                movel(spat_flatM_up_p, a=1.2, v=0.25, r=0.05)
                $ 2925 "Spatula_otw" "noBreak"
                movel(Spatula_otw_p, a=1.2, v=0.25)
                $ 2926 "switch_spat_F_M≔ False " "noBreak"
                global switch_spat_F_M=  False
              else:
                $ 2927 "ElseIf spatula≟'spatula_flat_S'" "noBreak"
                if (spatula == "spatula_flat_S"):
                  $ 2928 "MoveJ" "noBreak"
                  $ 2929 "Spatula_otw" "noBreak"
                  movej(get_inverse_kin(Spatula_otw_p, qnear=Spatula_otw_q), a=1.3962634015954636, v=1.0471975511965976)
                  $ 2930 "spat_flatS_up" "noBreak"
                  movej(get_inverse_kin(spat_flatS_up_p, qnear=spat_flatS_up_q), a=1.3962634015954636, v=1.0471975511965976, r=0.05)
                  $ 2931 "MoveL" "noBreak"
                  $ 2932 "spat_flatS_pick" "noBreak"
                  movel(spat_flatS_pick_p, a=1.2, v=0.25)
                  # begin: URCap Program Node
                  #   Source: Robotiq_Grippers, 3.17.0.105337, Robotiq Inc.
                  #   Type: Gripper
                  $ 2933 "Gripper Close (1)" "noBreak"
                  if not(gripper_connected[0]):
                    popup("Gripper 1 must be connected to run this program.", "No connection", False, True, True)
                  end
                  if not(rq_is_gripper_activated("1")):
                    popup("Gripper 1 is not activated. Go to Installation tab > Gripper to activate it and run the program again.", "Not activated", False, True, True)
                  end
                  rq_set_pos_spd_for(255, 0, 77, "1")
                  rq_wait_pos_spe_for_request(255, 0, 77, "1")
                  rq_go_to("1")
                  rq_wait("1")
                  # end: URCap Program Node
                  $ 2934 "spat_flatS_up" "noBreak"
                  movel(spat_flatS_up_p, a=1.2, v=0.25, r=0.05)
                  $ 2935 "Spatula_otw" "noBreak"
                  movel(Spatula_otw_p, a=1.2, v=0.25)
                  $ 2936 "switch_spat_F_S≔ False " "noBreak"
                  global switch_spat_F_S=  False
                end
              end
            end
          end
        end
        $ 2937 "weight_value≔get_weight()" "noBreak"
        global weight_value=get_weight()
        $ 2938 "auto_tilt_and_scoop(W_now, target_weight, weight_value)" "noBreak"
        auto_tilt_and_scoop(W_now, target_weight, weight_value)
        # begin: URCap Program Node
        #   Source: SensoPart VISOR Robotic, 2.0.6, SensoPart Industriesensorik GmbH
        #   Type: Approach Pose
        $ 2939 "Approach Pose" "noBreak"
        movej(pose_trans(easyPickPose,p[0.0000,0.0000,-0.0000,0.0000,0.0000,0.0000]),a=0.2618,v=0.1745,t=0.000000,r=0.000000)
        # end: URCap Program Node
        # begin: URCap Program Node
        #   Source: SensoPart VISOR Robotic, 2.0.6, SensoPart Industriesensorik GmbH
        #   Type: Target Pose
        $ 2940 "Target Pose" "noBreak"
        movel(pose_trans(easyPickPose,p[0.0000,0.0000,-0.0000,0.0000,0.0000,0.0000]),a=0.0500,v=0.0200,t=0.000000,r=0.000000)
        # end: URCap Program Node
        $ 2941 "Close Gripper" "noBreak"
        $ 2942 "dispense_pos≔get_actual_tcp_pose()" "noBreak"
        global dispense_pos= get_actual_tcp_pose ()
        $ 2943 "Loop weight_value≤target_weight" "noBreak"
        thread Thread_while_2943():
          while (True):
            $ 2944 "MoveL" "noBreak"
            $ 2945 "dispense_pos" "noBreak"
            movel(dispense_pos, a=0.2, v=0.1)
            $ 2946 "log_weight()" "noBreak"
            log_weight()
            $ 2947 "Wait: 0.5" "noBreak"
            sleep(0.5)
            $ 2948 "If level≥90.0" "noBreak"
            if (level >= 90.0):
              $ 2949 "Rotate()" "noBreak"
              Rotate()
            end
            $ 2950 "If level≤85" "noBreak"
            if (level <= 85):
              $ 2951 "tilt_to_home()" "noBreak"
              tilt_to_home()
            end
            $ 2952 "Wait: 0.5" "noBreak"
            sleep(0.5)
            $ 2953 "Start_thread≔ True " "noBreak"
            global Start_thread=  True
            $ 2954 "vib_thread≔ True " "noBreak"
            global vib_thread=  True
            $ 2956 "Wait: 0.5" "noBreak"
            sleep(0.5)
            $ 2962 "If diff ≥(target_g +(0.1*target_g))" "noBreak"
            if (diff  >= (target_g +(0.1*target_g))):
              $ 2963 "tilt_pose≔pose_trans(get_actual_tcp_pose(), p[0, 0, 0, 0, 0, 2.0])" "noBreak"
              global tilt_pose=pose_trans(get_actual_tcp_pose(), p[0, 0, 0, 0, 0, 2.0])
              $ 2964 "movel(tilt_pose, a=0.1, v=0.1, r=0.00001)" "noBreak"
              movel(tilt_pose, a=0.1, v=0.1, r=0.00001)
            else:
              $ 2965 "Else" "noBreak"
              $ 2966 "Loop weight_value≤target_weight and tilt_angle≥(-1.999) and tilt_angle≤0.5" "noBreak"
              thread Thread_while_2966():
                while (True):
                  $ 2967 "current_error≔target_weight-weight_value" "noBreak"
                  global current_error=target_weight-weight_value
                  $ 2968 "Integral_error≔Integral_error+current_error*dt" "noBreak"
                  global Integral_error=Integral_error+current_error*dt
                  $ 2969 "derivative≔(current_error-previous_error)/dt" "noBreak"
                  global derivative=(current_error-previous_error)/dt
                  $ 2970 "tilt_increment≔(kp*current_error)+(ki*Integral_error)+(kd*derivative)" "noBreak"
                  global tilt_increment=(kp*current_error)+(ki*Integral_error)+(kd*derivative)
                  $ 2971 "current_pose≔get_actual_tcp_pose()" "noBreak"
                  global current_pose= get_actual_tcp_pose ()
                  $ 2972 "tilt_angle≔current_pose[5]" "noBreak"
                  global tilt_angle=current_pose[5]
                  $ 2973 "tilt_pose≔pose_trans(current_pose, p[0, 0, 0, 0, 0, tilt_increment])" "noBreak"
                  global tilt_pose=pose_trans(current_pose, p[0, 0, 0, 0, 0, tilt_increment])
                  $ 2974 "movel(tilt_pose, a=0.1, v=0.1, r=0.00001)" "noBreak"
                  movel(tilt_pose, a=0.1, v=0.1, r=0.00001)
                  $ 2975 "previous_error≔current_error" "noBreak"
                  global previous_error=current_error
                end
              end
              if (weight_value <= target_weight  and  tilt_angle >= (-1.999)  and  tilt_angle <= 0.5):
                global thread_handler_2966=run Thread_while_2966()
                while (weight_value <= target_weight  and  tilt_angle >= (-1.999)  and  tilt_angle <= 0.5):
                  sync()
                end
                kill thread_handler_2966
              end
            end
            $ 2976 "Start_thread≔ False " "noBreak"
            global Start_thread=  False
            $ 2978 "weight_value≔get_weight()" "noBreak"
            global weight_value=get_weight()
            $ 2979 "tilt_angle≔-1" "noBreak"
            global tilt_angle=-1
            $ 2980 "Wait: 0.5" "noBreak"
            sleep(0.5)
            $ 2981 "vib_thread≔ False " "noBreak"
            global vib_thread=  False
            $ 2982 "MoveL" "noBreak"
            $ 2983 "dispense_pos" "noBreak"
            movel(dispense_pos, a=0.5, v=0.25)
            $ 2984 "compute_level_percent(W_now, weight_value)" "noBreak"
            compute_level_percent(W_now, weight_value)
            $ 2985 "send_level_info()" "noBreak"
            send_level_info()
            $ 2987 "spatula≔select_spatula(Flowability,level,diff,density)" "noBreak"
            global spatula=select_spatula(Flowability,level,diff,density)
            $ 2989 "Wait: 0.2" "noBreak"
            sleep(0.2)
            $ 2991 "Integral_error≔0" "noBreak"
            global Integral_error=0
            $ 2992 "current_error≔0" "noBreak"
            global current_error=0
            $ 2993 "previous_error≔0" "noBreak"
            global previous_error=0
            $ 2994 "Set AO[0]=0.0" "noBreak"
            set_standard_analog_out(0, 0.0)
            $ 2995 "Wait: 0.2" "noBreak"
            sleep(0.2)
            $ 2996 "send_spatula_info()" "noBreak"
            send_spatula_info()
            $ 2997 "If spatula ≟ 'spatula_M' and switch_spat_M≟ True " "noBreak"
            if (spatula  ==  "spatula_M"  and  switch_spat_M ==   True  ):
              $ 2998 "MoveJ" "noBreak"
              $ 2999 "Spatula_otw" "noBreak"
              movej(get_inverse_kin(Spatula_otw_p, qnear=Spatula_otw_q), a=1.3962634015954636, v=1.0471975511965976)
              $ 3000 "spat_L_up" "noBreak"
              movej(get_inverse_kin(spat_L_up_p, qnear=spat_L_up_q), a=1.3962634015954636, v=1.0471975511965976)
              $ 3001 "MoveL" "noBreak"
              $ 3002 "spat_L_side" "noBreak"
              movel(spat_L_side_p, a=1.2, v=0.25)
              $ 3003 "spat_L_lift" "noBreak"
              movel(spat_L_lift_p, a=1.2, v=0.25)
              $ 3004 "spat_L_pick" "noBreak"
              movel(spat_L_pick_p, a=1.2, v=0.25)
              # begin: URCap Program Node
              #   Source: Robotiq_Grippers, 3.17.0.105337, Robotiq Inc.
              #   Type: Gripper
              $ 3005 "Gripper Open (1)" "noBreak"
              if not(gripper_connected[0]):
                popup("Gripper 1 must be connected to run this program.", "No connection", False, True, True)
              end
              if not(rq_is_gripper_activated("1")):
                popup("Gripper 1 is not activated. Go to Installation tab > Gripper to activate it and run the program again.", "Not activated", False, True, True)
              end
              rq_set_pos_spd_for(0, 255, 77, "1")
              rq_wait_pos_spe_for_request(0, 255, 77, "1")
              rq_go_to("1")
              rq_wait("1")
              # end: URCap Program Node
              $ 3006 "spat_M_pick" "noBreak"
              movel(spat_M_pick_p, a=1.2, v=0.25)
              # begin: URCap Program Node
              #   Source: Robotiq_Grippers, 3.17.0.105337, Robotiq Inc.
              #   Type: Gripper
              $ 3007 "Gripper Close (1)" "noBreak"
              if not(gripper_connected[0]):
                popup("Gripper 1 must be connected to run this program.", "No connection", False, True, True)
              end
              if not(rq_is_gripper_activated("1")):
                popup("Gripper 1 is not activated. Go to Installation tab > Gripper to activate it and run the program again.", "Not activated", False, True, True)
              end
              rq_set_pos_spd_for(255, 0, 77, "1")
              rq_wait_pos_spe_for_request(255, 0, 77, "1")
              rq_go_to("1")
              rq_wait("1")
              # end: URCap Program Node
              $ 3008 "spat_M_up" "noBreak"
              movel(spat_M_up_p, a=1.2, v=0.25)
              $ 3009 "Spatula_otw" "noBreak"
              movel(Spatula_otw_p, a=1.2, v=0.25)
              $ 3010 "switch_spat_M≔ False " "noBreak"
              global switch_spat_M=  False
            else:
              $ 3011 "ElseIf spatula ≟ 'spatula_S' and switch_spat_S ≟ True " "noBreak"
              if (spatula  ==  "spatula_S" and switch_spat_S  ==   True  ):
                $ 3012 "MoveL" "noBreak"
                $ 3013 "Spatula_otw" "noBreak"
                movel(Spatula_otw_p, a=1.2, v=0.25)
                $ 3014 "spat_M_up" "noBreak"
                movel(spat_M_up_p, a=1.2, v=0.25)
                $ 3015 "spat_M_pick" "noBreak"
                movel(spat_M_pick_p, a=1.2, v=0.25)
                # begin: URCap Program Node
                #   Source: Robotiq_Grippers, 3.17.0.105337, Robotiq Inc.
                #   Type: Gripper
                $ 3016 "Gripper Open (1)" "noBreak"
                if not(gripper_connected[0]):
                  popup("Gripper 1 must be connected to run this program.", "No connection", False, True, True)
                end
                if not(rq_is_gripper_activated("1")):
                  popup("Gripper 1 is not activated. Go to Installation tab > Gripper to activate it and run the program again.", "Not activated", False, True, True)
                end
                rq_set_pos_spd_for(0, 255, 77, "1")
                rq_wait_pos_spe_for_request(0, 255, 77, "1")
                rq_go_to("1")
                rq_wait("1")
                # end: URCap Program Node
                $ 3017 "spat_S_pick" "noBreak"
                movel(spat_S_pick_p, a=1.2, v=0.25)
                # begin: URCap Program Node
                #   Source: Robotiq_Grippers, 3.17.0.105337, Robotiq Inc.
                #   Type: Gripper
                $ 3018 "Gripper Close (1)" "noBreak"
                if not(gripper_connected[0]):
                  popup("Gripper 1 must be connected to run this program.", "No connection", False, True, True)
                end
                if not(rq_is_gripper_activated("1")):
                  popup("Gripper 1 is not activated. Go to Installation tab > Gripper to activate it and run the program again.", "Not activated", False, True, True)
                end
                rq_set_pos_spd_for(255, 0, 77, "1")
                rq_wait_pos_spe_for_request(255, 0, 77, "1")
                rq_go_to("1")
                rq_wait("1")
                # end: URCap Program Node
                $ 3019 "spat_S_up" "noBreak"
                movel(spat_S_up_p, a=1.2, v=0.25)
                $ 3020 "Spatula_otw" "noBreak"
                movel(Spatula_otw_p, a=1.2, v=0.25)
                $ 3021 "switch_spat_S≔ False " "noBreak"
                global switch_spat_S=  False
              else:
                $ 3022 "ElseIf spatula≟'spatula_flat_S'  and switch_spat_F_S ≟ True " "noBreak"
                if (spatula == "spatula_flat_S"   and  switch_spat_F_S  ==   True  ):
                  $ 3023 "MoveL" "noBreak"
                  $ 3024 "Spatula_otw" "noBreak"
                  movel(Spatula_otw_p, a=1.2, v=0.25)
                  $ 3025 "spat_flatM_up" "noBreak"
                  movel(spat_flatM_up_p, a=1.2, v=0.25)
                  $ 3026 "spat_flatM_pick" "noBreak"
                  movel(spat_flatM_pick_p, a=1.2, v=0.25)
                  # begin: URCap Program Node
                  #   Source: Robotiq_Grippers, 3.17.0.105337, Robotiq Inc.
                  #   Type: Gripper
                  $ 3027 "Gripper Open (1)" "noBreak"
                  if not(gripper_connected[0]):
                    popup("Gripper 1 must be connected to run this program.", "No connection", False, True, True)
                  end
                  if not(rq_is_gripper_activated("1")):
                    popup("Gripper 1 is not activated. Go to Installation tab > Gripper to activate it and run the program again.", "Not activated", False, True, True)
                  end
                  rq_set_pos_spd_for(0, 0, 77, "1")
                  rq_wait_pos_spe_for_request(0, 0, 77, "1")
                  rq_go_to("1")
                  rq_wait("1")
                  # end: URCap Program Node
                  $ 3028 "spat_flatS_pick" "noBreak"
                  movel(spat_flatS_pick_p, a=1.2, v=0.25)
                  # begin: URCap Program Node
                  #   Source: Robotiq_Grippers, 3.17.0.105337, Robotiq Inc.
                  #   Type: Gripper
                  $ 3029 "Gripper Close (1)" "noBreak"
                  if not(gripper_connected[0]):
                    popup("Gripper 1 must be connected to run this program.", "No connection", False, True, True)
                  end
                  if not(rq_is_gripper_activated("1")):
                    popup("Gripper 1 is not activated. Go to Installation tab > Gripper to activate it and run the program again.", "Not activated", False, True, True)
                  end
                  rq_set_pos_spd_for(255, 0, 77, "1")
                  rq_wait_pos_spe_for_request(255, 0, 77, "1")
                  rq_go_to("1")
                  rq_wait("1")
                  # end: URCap Program Node
                  $ 3030 "spat_flatS_up" "noBreak"
                  movel(spat_flatS_up_p, a=1.2, v=0.25)
                  $ 3031 "Spatula_otw" "noBreak"
                  movel(Spatula_otw_p, a=1.2, v=0.25)
                  $ 3032 "switch_spat_F_S≔ False " "noBreak"
                  global switch_spat_F_S=  False
                end
              end
            end
            $ 3033 "auto_tilt_and_scoop(W_now, target_weight, weight_value)" "noBreak"
            auto_tilt_and_scoop(W_now, target_weight, weight_value)
            $ 3034 "Wait: 0.5" "noBreak"
            sleep(0.5)
          end
        end
        if (weight_value <= target_weight):
          global thread_handler_2943=run Thread_while_2943()
          while (weight_value <= target_weight):
            sync()
          end
          kill thread_handler_2943
        end
        $ 3035 "Start_thread≔ False " "noBreak"
        global Start_thread=  False
        $ 3036 "Wait: 0.5" "noBreak"
        sleep(0.5)
        $ 3037 "vib_thread≔ False " "noBreak"
        global vib_thread=  False
        # begin: URCap Program Node
        #   Source: SensoPart VISOR Robotic, 2.0.6, SensoPart Industriesensorik GmbH
        #   Type: Exit Pose
        $ 3039 "Exit Pose" "noBreak"
        movel(pose_trans(easyPickPose,p[0.0000,0.0000,-0.0000,0.0000,0.0000,0.0000]),a=0.5000,v=0.2500,t=0.000000,r=0.000000)
        # end: URCap Program Node
        easyPickObjTaken = True
      end
      # end: URCap Program Node
      # begin: URCap Program Node
      #   Source: SensoPart VISOR Robotic, 2.0.6, SensoPart Industriesensorik GmbH
      #   Type: No Object Detected
      $ 3040 "No Object Detected" "noBreak"
      if (visor_partsFound(easyPickVisorId) < 1):
        $ 3041 "Popup: No weigh scale detected" "noBreak"
        popup("No weigh scale detected", "Message", False, False, blocking=True)
        else:
      end
      # end: URCap Program Node
    end
    easyPickCount_4 = easyPickCount_4 + 1
    visor_easyPickUpdate(easyPickVisorId, "counter", easyPickCount_4)
    visor_easyPickSetIdent("6c09fd", easyPickVisorId)
    # end: URCap Program Node
  end
  visorFuncEasyPick_ff2f00()
  # end: URCap Program Node
  $ 3044 "MoveJ"
  $ 3045 "dispense_pos" "breakAfter"
  movej(dispense_pos, a=0.5235987755982988, v=0.4363323129985824)
  $ 3046 "after_scoop()"
  after_scoop()
  $ 3047 "Place spatula back to the rack"
  $ 3048 "If spatula≟'spatula_M'"
  if (spatula == "spatula_M"):
    $ 3049 "MoveJ"
    $ 3050 "Spatula_otw" "breakAfter"
    movej(get_inverse_kin(Spatula_otw_p, qnear=Spatula_otw_q), a=1.3962634015954636, v=1.0471975511965976)
    $ 3051 "spat_M_up" "breakAfter"
    movej(get_inverse_kin(spat_M_up_p, qnear=spat_M_up_q), a=1.3962634015954636, v=1.0471975511965976)
    $ 3052 "MoveL"
    $ 3053 "spat_M_pick" "breakAfter"
    movel(spat_M_pick_p, a=1.2, v=0.25)
    # begin: URCap Program Node
    #   Source: Robotiq_Grippers, 3.17.0.105337, Robotiq Inc.
    #   Type: Gripper
    $ 3054 "Gripper Open (1)"
    if not(gripper_connected[0]):
      popup("Gripper 1 must be connected to run this program.", "No connection", False, True, True)
    end
    if not(rq_is_gripper_activated("1")):
      popup("Gripper 1 is not activated. Go to Installation tab > Gripper to activate it and run the program again.", "Not activated", False, True, True)
    end
    rq_set_pos_spd_for(0, 128, 77, "1")
    rq_wait_pos_spe_for_request(0, 128, 77, "1")
    rq_go_to("1")
    rq_wait("1")
    # end: URCap Program Node
    $ 3055 "spat_M_up" "breakAfter"
    movel(spat_M_up_p, a=1.2, v=0.25)
    $ 3056 "Home (Safe)"
    movej([-1.2302089344500047, -1.2969853503591224, -1.875639182904262, -1.539621866126728, 1.5731943360401213, -2.80099559440227], a=1.3962634015954636, v=1.0471975511965976)
  else:
    $ 3057 "ElseIf spatula≟'spatula_flat_S'"
    if (spatula == "spatula_flat_S"):
      $ 3058 "MoveJ"
      $ 3059 "Spatula_otw" "breakAfter"
      movej(get_inverse_kin(Spatula_otw_p, qnear=Spatula_otw_q), a=1.3962634015954636, v=1.0471975511965976)
      $ 3060 "spat_flatS_up" "breakAfter"
      movej(get_inverse_kin(spat_flatS_up_p, qnear=spat_flatS_up_q), a=1.3962634015954636, v=1.0471975511965976)
      $ 3061 "MoveL"
      $ 3062 "spat_flatS_pick" "breakAfter"
      movel(spat_flatS_pick_p, a=1.2, v=0.25)
      # begin: URCap Program Node
      #   Source: Robotiq_Grippers, 3.17.0.105337, Robotiq Inc.
      #   Type: Gripper
      $ 3063 "Gripper Open (1)"
      if not(gripper_connected[0]):
        popup("Gripper 1 must be connected to run this program.", "No connection", False, True, True)
      end
      if not(rq_is_gripper_activated("1")):
        popup("Gripper 1 is not activated. Go to Installation tab > Gripper to activate it and run the program again.", "Not activated", False, True, True)
      end
      rq_set_pos_spd_for(0, 128, 77, "1")
      rq_wait_pos_spe_for_request(0, 128, 77, "1")
      rq_go_to("1")
      rq_wait("1")
      # end: URCap Program Node
      $ 3064 "spat_flatS_up" "breakAfter"
      movel(spat_flatS_up_p, a=1.2, v=0.25)
      $ 3065 "Home (Safe)"
      movej([-1.2302089344500047, -1.2969853503591224, -1.875639182904262, -1.539621866126728, 1.5731943360401213, -2.80099559440227], a=1.3962634015954636, v=1.0471975511965976)
    end
  end
  $ 3066 "Pick container from PoTS"
  $ 3067 "cont_place_offs≔pose_add(container_place, p[0.05,0,0,0,0,0])"
  global cont_place_offs=pose_add(container_place, p[0.05,0,0,0,0,0])
  $ 3068 "MoveJ"
  $ 3069 "cont_place_offs" "breakAfter"
  movej(cont_place_offs, a=1.3962634015954636, v=1.0471975511965976)
  $ 3070 "container_place" "breakAfter"
  movej(container_place, a=1.3962634015954636, v=1.0471975511965976)
  $ 3071 "MoveL"
  $ 3072 "target_pose" "breakAfter"
  movel(target_pose, a=1.2, v=0.25)
  # begin: URCap Program Node
  #   Source: Robotiq_Grippers, 3.17.0.105337, Robotiq Inc.
  #   Type: Gripper
  $ 3073 "Gripper Close (1)"
  if not(gripper_connected[0]):
    popup("Gripper 1 must be connected to run this program.", "No connection", False, True, True)
  end
  if not(rq_is_gripper_activated("1")):
    popup("Gripper 1 is not activated. Go to Installation tab > Gripper to activate it and run the program again.", "Not activated", False, True, True)
  end
  rq_set_pos_spd_for(255, 77, 77, "1")
  rq_wait_pos_spe_for_request(255, 77, 77, "1")
  rq_go_to("1")
  rq_wait("1")
  # end: URCap Program Node
  $ 3074 "container_place" "breakAfter"
  movel(container_place, a=0.6, v=0.1)
  $ 3075 "powder_position≔'Position1'"
  global powder_position="Position1"
  $ 3076 "Place Powder container back to holder"
  $ 3077 "If powder_position ≟ 'Position1'"
  if (powder_position  ==  "Position1"):
    $ 3078 "MoveL"
    $ 3079 "Postions_otw" "breakAfter"
    movel(Postions_otw_p, a=1.2, v=0.25, r=0.01)
    $ 3080 "MoveL"
    $ 3081 "PosA_up" "breakAfter"
    movel(PosA_up_p, a=1.2, v=0.25)
    $ 3082 "PosA_pick" "breakAfter"
    movel(PosA_pick_p, a=0.3, v=0.05)
    # begin: URCap Program Node
    #   Source: Robotiq_Grippers, 3.17.0.105337, Robotiq Inc.
    #   Type: Gripper
    $ 3083 "Gripper Open (1)"
    if not(gripper_connected[0]):
      popup("Gripper 1 must be connected to run this program.", "No connection", False, True, True)
    end
    if not(rq_is_gripper_activated("1")):
      popup("Gripper 1 is not activated. Go to Installation tab > Gripper to activate it and run the program again.", "Not activated", False, True, True)
    end
    rq_set_pos_spd_for(0, 128, 77, "1")
    rq_wait_pos_spe_for_request(0, 128, 77, "1")
    rq_go_to("1")
    rq_wait("1")
    # end: URCap Program Node
    $ 3084 "PosA_up" "breakAfter"
    movel(PosA_up_p, a=1.2, v=0.25)
    $ 3085 "Postions_otw" "breakAfter"
    movel(Postions_otw_p, a=1.2, v=0.25, r=0.05)
  else:
    $ 3086 "ElseIf powder_position≟'Position2'"
    if (powder_position == "Position2"):
      $ 3087 "MoveL"
      $ 3088 "Postions_otw" "breakAfter"
      movel(Postions_otw_p, a=1.2, v=0.25, r=0.01)
      $ 3089 "MoveL"
      $ 3090 "PosB_up" "breakAfter"
      movel(PosB_up_p, a=1.2, v=0.25, r=0.01)
      $ 3091 "PosB_pick" "breakAfter"
      movel(PosB_pick_p, a=0.3, v=0.05)
      # begin: URCap Program Node
      #   Source: Robotiq_Grippers, 3.17.0.105337, Robotiq Inc.
      #   Type: Gripper
      $ 3092 "Gripper Open (1)"
      if not(gripper_connected[0]):
        popup("Gripper 1 must be connected to run this program.", "No connection", False, True, True)
      end
      if not(rq_is_gripper_activated("1")):
        popup("Gripper 1 is not activated. Go to Installation tab > Gripper to activate it and run the program again.", "Not activated", False, True, True)
      end
      rq_set_pos_spd_for(0, 128, 77, "1")
      rq_wait_pos_spe_for_request(0, 128, 77, "1")
      rq_go_to("1")
      rq_wait("1")
      # end: URCap Program Node
      $ 3093 "PosB_up" "breakAfter"
      movel(PosB_up_p, a=1.2, v=0.25)
      $ 3094 "Postions_otw" "breakAfter"
      movel(Postions_otw_p, a=1.2, v=0.25, r=0.05)
    else:
      $ 3095 "ElseIf powder_position≟'Position3'"
      if (powder_position == "Position3"):
        $ 3096 "MoveL"
        $ 3097 "Postions_otw" "breakAfter"
        movel(Postions_otw_p, a=1.2, v=0.25, r=0.01)
        $ 3098 "MoveL"
        $ 3099 "PosC_up" "breakAfter"
        movel(PosC_up_p, a=1.2, v=0.25, r=0.01)
        $ 3100 "PosC_pick" "breakAfter"
        movel(PosC_pick_p, a=0.3, v=0.05)
        # begin: URCap Program Node
        #   Source: Robotiq_Grippers, 3.17.0.105337, Robotiq Inc.
        #   Type: Gripper
        $ 3101 "Gripper Open (1)"
        if not(gripper_connected[0]):
          popup("Gripper 1 must be connected to run this program.", "No connection", False, True, True)
        end
        if not(rq_is_gripper_activated("1")):
          popup("Gripper 1 is not activated. Go to Installation tab > Gripper to activate it and run the program again.", "Not activated", False, True, True)
        end
        rq_set_pos_spd_for(0, 128, 77, "1")
        rq_wait_pos_spe_for_request(0, 128, 77, "1")
        rq_go_to("1")
        rq_wait("1")
        # end: URCap Program Node
        $ 3102 "PosC_up" "breakAfter"
        movel(PosC_up_p, a=1.2, v=0.25)
        $ 3103 "Postions_otw" "breakAfter"
        movel(Postions_otw_p, a=1.2, v=0.25, r=0.05)
      end
    end
  end
  $ 3104 "Cap the container"
  $ 3105 "If powder_position ≟ 'Position1'"
  if (powder_position  ==  "Position1"):
    $ 3106 "MoveJ"
    $ 3107 "Cap_Pos1_up" "breakAfter"
    movej(get_inverse_kin(Cap_Pos1_up_p, qnear=Cap_Pos1_up_q), a=1.3962634015954636, v=1.0471975511965976)
    $ 3108 "MoveL"
    $ 3109 "Cap_pos1" "breakAfter"
    movel(Cap_pos1_p, a=0.3, v=0.05)
  else:
    $ 3110 "ElseIf powder_position≟'Position2'"
    if (powder_position == "Position2"):
      $ 3111 "MoveJ"
      $ 3112 "Cap_Pos2_up" "breakAfter"
      movej(get_inverse_kin(Cap_Pos2_up_p, qnear=Cap_Pos2_up_q), a=1.3962634015954636, v=1.0471975511965976)
      $ 3113 "MoveL"
      $ 3114 "Cap_Pos2" "breakAfter"
      movel(Cap_Pos2_p, a=0.3, v=0.05)
    else:
      $ 3115 "ElseIf powder_position≟'Position3'"
      if (powder_position == "Position3"):
        $ 3116 "MoveJ"
        $ 3117 "Cap_Pos3_up" "breakAfter"
        movej(get_inverse_kin(Cap_Pos3_up_p, qnear=Cap_Pos3_up_q), a=1.3962634015954636, v=1.0471975511965976)
        $ 3118 "MoveL"
        $ 3119 "Cap_pos3" "breakAfter"
        movel(Cap_pos3_p, a=0.3, v=0.05)
      end
    end
  end
  $ 3120 "Capping motion"
  # begin: URCap Program Node
  #   Source: Robotiq_Grippers, 3.17.0.105337, Robotiq Inc.
  #   Type: Gripper
  $ 3121 "Gripper Move30mm (1)"
  if not(gripper_connected[0]):
    popup("Gripper 1 must be connected to run this program.", "No connection", False, True, True)
  end
  if not(rq_is_gripper_activated("1")):
    popup("Gripper 1 is not activated. Go to Installation tab > Gripper to activate it and run the program again.", "Not activated", False, True, True)
  end
  rq_set_pos_spd_for(110, 77, 77, "1")
  rq_wait_pos_spe_for_request(110, 77, 77, "1")
  rq_go_to("1")
  rq_wait("1")
  # end: URCap Program Node
  $ 3122 "Loop 2 times"
  Loop_4 = 0
  while (Loop_4 < 2):
    $ 3128 "Cap_CW≔pose_add(get_actual_tcp_pose(), p[0,0,0,0,0,2.2])"
    global Cap_CW= pose_add ( get_actual_tcp_pose (), p[0,0,0,0,0,2.2])
    $ 3129 "MoveL"
    $ 3130 "Cap_CW" "breakAfter"
    movel(Cap_CW, a=1.2, v=0.25)
    # begin: URCap Program Node
    #   Source: Robotiq_Grippers, 3.17.0.105337, Robotiq Inc.
    #   Type: Gripper
    $ 3131 "Gripper Move25mm (1)"
    if not(gripper_connected[0]):
      popup("Gripper 1 must be connected to run this program.", "No connection", False, True, True)
    end
    if not(rq_is_gripper_activated("1")):
      popup("Gripper 1 is not activated. Go to Installation tab > Gripper to activate it and run the program again.", "Not activated", False, True, True)
    end
    rq_set_pos_spd_for(133, 77, 77, "1")
    rq_wait_pos_spe_for_request(133, 77, 77, "1")
    rq_go_to("1")
    rq_wait("1")
    # end: URCap Program Node
    $ 3132 "Cap_CCW≔pose_add(get_actual_tcp_pose(), p[0,0,0,0,0,-2.2])"
    global Cap_CCW= pose_add ( get_actual_tcp_pose (), p[0,0,0,0,0,-2.2])
    $ 3133 "MoveL"
    $ 3134 "Cap_CCW" "breakAfter"
    movel(Cap_CCW, a=1.2, v=0.25)
    # begin: URCap Program Node
    #   Source: Robotiq_Grippers, 3.17.0.105337, Robotiq Inc.
    #   Type: Gripper
    $ 3135 "Gripper Move30mm (1)"
    if not(gripper_connected[0]):
      popup("Gripper 1 must be connected to run this program.", "No connection", False, True, True)
    end
    if not(rq_is_gripper_activated("1")):
      popup("Gripper 1 is not activated. Go to Installation tab > Gripper to activate it and run the program again.", "Not activated", False, True, True)
    end
    rq_set_pos_spd_for(110, 77, 77, "1")
    rq_wait_pos_spe_for_request(110, 77, 77, "1")
    rq_go_to("1")
    rq_wait("1")
    # end: URCap Program Node
    Loop_4 = Loop_4 + 1
  end
  # begin: URCap Program Node
  #   Source: Robotiq_Grippers, 3.17.0.105337, Robotiq Inc.
  #   Type: Gripper
  $ 3136 "Gripper Open (1)"
  if not(gripper_connected[0]):
    popup("Gripper 1 must be connected to run this program.", "No connection", False, True, True)
  end
  if not(rq_is_gripper_activated("1")):
    popup("Gripper 1 is not activated. Go to Installation tab > Gripper to activate it and run the program again.", "Not activated", False, True, True)
  end
  rq_set_pos_spd_for(0, 77, 77, "1")
  rq_wait_pos_spe_for_request(0, 77, 77, "1")
  rq_go_to("1")
  rq_wait("1")
  # end: URCap Program Node
  $ 3137 "after_capping≔pose_add(get_actual_tcp_pose(), p[0,0,0.05,0,0,0])"
  global after_capping=pose_add(get_actual_tcp_pose(), p[0,0,0.05,0,0,0])
  $ 3138 "MoveL"
  $ 3139 "after_capping" "breakAfter"
  movel(after_capping, a=1.2, v=0.25)
  $ 3140 "Home (Safe)"
  movej([-1.2302089344500047, -1.2969853503591224, -1.875639182904262, -1.539621866126728, 1.5731943360401213, -2.80099559440227], a=1.3962634015954636, v=1.0471975511965976)
  elif (44 == switch_1):
    $ 3203 "Case 44"
    $ 3204 "Decap Container for recipe"
    $ 3206 "If powder_position ≟ 'Position1'"
    if (powder_position  ==  "Position1"):
      $ 3207 "MoveJ"
      $ 3208 "Postions_otw" "breakAfter"
      movej(get_inverse_kin(Postions_otw_p, qnear=Postions_otw_q), a=1.3962634015954636, v=1.0471975511965976, r=0.01)
      # begin: URCap Program Node
      #   Source: Robotiq_Grippers, 3.17.0.105337, Robotiq Inc.
      #   Type: Gripper
      $ 3209 "Gripper Open (1)"
      if not(gripper_connected[0]):
        popup("Gripper 1 must be connected to run this program.", "No connection", False, True, True)
      end
      if not(rq_is_gripper_activated("1")):
        popup("Gripper 1 is not activated. Go to Installation tab > Gripper to activate it and run the program again.", "Not activated", False, True, True)
      end
      rq_set_pos_spd_for(0, 127, 77, "1")
      rq_wait_pos_spe_for_request(0, 127, 77, "1")
      rq_go_to("1")
      rq_wait("1")
      # end: URCap Program Node
      $ 3210 "MoveL"
      $ 3211 "PosA_up" "breakAfter"
      movel(PosA_up_p, a=1.2, v=0.25)
      $ 3212 "PosA_pick" "breakAfter"
      movel(PosA_pick_p, a=1.2, v=0.25)
      # begin: URCap Program Node
      #   Source: Robotiq_Grippers, 3.17.0.105337, Robotiq Inc.
      #   Type: Gripper
      $ 3213 "Gripper Close (1)"
      if not(gripper_connected[0]):
        popup("Gripper 1 must be connected to run this program.", "No connection", False, True, True)
      end
      if not(rq_is_gripper_activated("1")):
        popup("Gripper 1 is not activated. Go to Installation tab > Gripper to activate it and run the program again.", "Not activated", False, True, True)
      end
      rq_set_pos_spd_for(255, 127, 77, "1")
      rq_wait_pos_spe_for_request(255, 127, 77, "1")
      rq_go_to("1")
      rq_wait("1")
      # end: URCap Program Node
      $ 3214 "PosA_up" "breakAfter"
      movel(PosA_up_p, a=0.3, v=0.04)
      $ 3215 "Postions_otw" "breakAfter"
      movel(Postions_otw_p, a=1.2, v=0.25, r=0.01)
    else:
      $ 3216 "ElseIf powder_position≟'Position2'"
      if (powder_position == "Position2"):
        $ 3217 "MoveJ"
        $ 3218 "Postions_otw" "breakAfter"
        movej(get_inverse_kin(Postions_otw_p, qnear=Postions_otw_q), a=1.3962634015954636, v=1.0471975511965976, r=0.01)
        # begin: URCap Program Node
        #   Source: Robotiq_Grippers, 3.17.0.105337, Robotiq Inc.
        #   Type: Gripper
        $ 3219 "Gripper Open (1)"
        if not(gripper_connected[0]):
          popup("Gripper 1 must be connected to run this program.", "No connection", False, True, True)
        end
        if not(rq_is_gripper_activated("1")):
          popup("Gripper 1 is not activated. Go to Installation tab > Gripper to activate it and run the program again.", "Not activated", False, True, True)
        end
        rq_set_pos_spd_for(0, 127, 77, "1")
        rq_wait_pos_spe_for_request(0, 127, 77, "1")
        rq_go_to("1")
        rq_wait("1")
        # end: URCap Program Node
        $ 3220 "MoveL"
        $ 3221 "PosB_up" "breakAfter"
        movel(PosB_up_p, a=1.2, v=0.25, r=0.01)
        $ 3222 "PosB_pick" "breakAfter"
        movel(PosB_pick_p, a=1.2, v=0.25)
        # begin: URCap Program Node
        #   Source: Robotiq_Grippers, 3.17.0.105337, Robotiq Inc.
        #   Type: Gripper
        $ 3223 "Gripper Close (1)"
        if not(gripper_connected[0]):
          popup("Gripper 1 must be connected to run this program.", "No connection", False, True, True)
        end
        if not(rq_is_gripper_activated("1")):
          popup("Gripper 1 is not activated. Go to Installation tab > Gripper to activate it and run the program again.", "Not activated", False, True, True)
        end
        rq_set_pos_spd_for(255, 127, 77, "1")
        rq_wait_pos_spe_for_request(255, 127, 77, "1")
        rq_go_to("1")
        rq_wait("1")
        # end: URCap Program Node
        $ 3224 "PosB_up" "breakAfter"
        movel(PosB_up_p, a=0.4, v=0.05)
        $ 3225 "Postions_otw" "breakAfter"
        movel(Postions_otw_p, a=1.2, v=0.25)
      else:
        $ 3226 "ElseIf powder_position≟'Position3'"
        if (powder_position == "Position3"):
          $ 3227 "MoveJ"
          $ 3228 "Postions_otw" "breakAfter"
          movej(get_inverse_kin(Postions_otw_p, qnear=Postions_otw_q), a=1.3962634015954636, v=1.0471975511965976, r=0.01)
          # begin: URCap Program Node
          #   Source: Robotiq_Grippers, 3.17.0.105337, Robotiq Inc.
          #   Type: Gripper
          $ 3229 "Gripper Open (1)"
          if not(gripper_connected[0]):
            popup("Gripper 1 must be connected to run this program.", "No connection", False, True, True)
          end
          if not(rq_is_gripper_activated("1")):
            popup("Gripper 1 is not activated. Go to Installation tab > Gripper to activate it and run the program again.", "Not activated", False, True, True)
          end
          rq_set_pos_spd_for(0, 127, 77, "1")
          rq_wait_pos_spe_for_request(0, 127, 77, "1")
          rq_go_to("1")
          rq_wait("1")
          # end: URCap Program Node
          $ 3230 "MoveL"
          $ 3231 "PosC_up" "breakAfter"
          movel(PosC_up_p, a=1.2, v=0.25, r=0.01)
          $ 3232 "PosC_pick" "breakAfter"
          movel(PosC_pick_p, a=1.2, v=0.25)
          # begin: URCap Program Node
          #   Source: Robotiq_Grippers, 3.17.0.105337, Robotiq Inc.
          #   Type: Gripper
          $ 3233 "Gripper Close (1)"
          if not(gripper_connected[0]):
            popup("Gripper 1 must be connected to run this program.", "No connection", False, True, True)
          end
          if not(rq_is_gripper_activated("1")):
            popup("Gripper 1 is not activated. Go to Installation tab > Gripper to activate it and run the program again.", "Not activated", False, True, True)
          end
          rq_set_pos_spd_for(255, 127, 77, "1")
          rq_wait_pos_spe_for_request(255, 127, 77, "1")
          rq_go_to("1")
          rq_wait("1")
          # end: URCap Program Node
          $ 3234 "PosC_up" "breakAfter"
          movel(PosC_up_p, a=0.5, v=0.05)
        end
      end
    end
    $ 3235 "MoveJ"
    $ 3236 "Pow_decap_up" "breakAfter"
    movej(get_inverse_kin(Pow_decap_up_p, qnear=Pow_decap_up_q), a=1.3962634015954636, v=1.0471975511965976)
    $ 3237 "Set GRP_3F_Open=On"
    set_standard_digital_out(5, True)
    $ 3238 "Wait: 0.5"
    sleep(0.5)
    $ 3239 "MoveL"
    $ 3240 "pow_decap_place" "breakAfter"
    movel(pow_decap_place_p, a=0.5, v=0.05)
    $ 3241 "Set GRP_3F_Open=Off"
    set_standard_digital_out(5, False)
    $ 3242 "Wait: 0.5"
    sleep(0.5)
    # begin: URCap Program Node
    #   Source: Robotiq_Grippers, 3.17.0.105337, Robotiq Inc.
    #   Type: Gripper
    $ 3243 "Gripper Open (1)"
    if not(gripper_connected[0]):
      popup("Gripper 1 must be connected to run this program.", "No connection", False, True, True)
    end
    if not(rq_is_gripper_activated("1")):
      popup("Gripper 1 is not activated. Go to Installation tab > Gripper to activate it and run the program again.", "Not activated", False, True, True)
    end
    rq_set_pos_spd_for(0, 255, 77, "1")
    rq_wait_pos_spe_for_request(0, 255, 77, "1")
    rq_go_to("1")
    rq_wait("1")
    # end: URCap Program Node
    $ 3244 "MoveL"
    $ 3245 "Pow_decap_up" "breakAfter"
    movel(Pow_decap_up_p, a=1.2, v=0.25)
    $ 3246 "Postions_otw" "breakAfter"
    movel(Postions_otw_p, a=1.2, v=0.25)
    $ 3247 "Home (Safe)"
    movej([-1.2302089344500047, -1.2969853503591224, -1.875639182904262, -1.539621866126728, 1.5731943360401213, -2.80099559440227], a=1.3962634015954636, v=1.0471975511965976)
    $ 3248 "MoveL"
    $ 3249 "Decap_above" "breakAfter"
    movel(Decap_above_p, a=1.2, v=0.25)
    $ 3250 "Decapp" "breakAfter"
    movel(Decapp_p, a=1.2, v=0.25)
    # begin: URCap Program Node
    #   Source: Robotiq_Grippers, 3.17.0.105337, Robotiq Inc.
    #   Type: Gripper
    $ 3251 "Gripper Close (1)"
    if not(gripper_connected[0]):
      popup("Gripper 1 must be connected to run this program.", "No connection", False, True, True)
    end
    if not(rq_is_gripper_activated("1")):
      popup("Gripper 1 is not activated. Go to Installation tab > Gripper to activate it and run the program again.", "Not activated", False, True, True)
    end
    rq_set_pos_spd_for(255, 128, 77, "1")
    rq_wait_pos_spe_for_request(255, 128, 77, "1")
    rq_go_to("1")
    rq_wait("1")
    # end: URCap Program Node
    $ 3252 "Decap"
    $ 3253 "Action_Info≔'decapping'"
    global Action_Info="decapping"
    $ 3254 "Set GRP_3F_Enable=On"
    set_standard_digital_out(4, True)
    $ 3255 "Set GRP_3F_Decap=On"
    set_standard_digital_out(3, True)
    $ 3256 "Force"
    sleep(0.02)
    zero_ftsensor()
    force_mode(p[0.0,0.0,0.0,0.0,0.0,0.0], [0, 0, 1, 0, 0, 0], [0.0, 0.0, 2.0, 0.0, 0.0, 0.0], 2, [0.1, 0.1, 5.0E-4, 0.3490658503988659, 0.3490658503988659, 0.3490658503988659])
    $ 3257 "check_decapping(offset=0.010, timeout=4.5, abort=CMD_Hold)" "noBreak"
    check_decapping(offset=0.010, timeout=4.5, abort=CMD_Hold)
    end_force_mode()
    stopl(5.0)
    $ 3258 "Set GRP_3F_Decap=Off"
    set_standard_digital_out(3, False)
    $ 3259 "Set GRP_3F_Enable=Off"
    set_standard_digital_out(4, False)
    $ 3260 "MoveL"
    $ 3261 "Decap_above" "breakAfter"
    movel(Decap_above_p, a=1.2, v=0.25)
    $ 3262 "Cap_above" "breakAfter"
    movel(Cap_above_p, a=1.2, v=0.25, r=0.05)
    $ 3263 "Cap_place" "breakAfter"
    movel(Cap_place_p, a=1.2, v=0.25)
    # begin: URCap Program Node
    #   Source: Robotiq_Grippers, 3.17.0.105337, Robotiq Inc.
    #   Type: Gripper
    $ 3264 "Gripper Move39mm (1)"
    if not(gripper_connected[0]):
      popup("Gripper 1 must be connected to run this program.", "No connection", False, True, True)
    end
    if not(rq_is_gripper_activated("1")):
      popup("Gripper 1 is not activated. Go to Installation tab > Gripper to activate it and run the program again.", "Not activated", False, True, True)
    end
    rq_set_pos_spd_for(67, 77, 77, "1")
    rq_wait_pos_spe_for_request(67, 77, 77, "1")
    rq_go_to("1")
    rq_wait("1")
    # end: URCap Program Node
    $ 3265 "Cap_above" "breakAfter"
    movel(Cap_above_p, a=1.2, v=0.25, r=0.05)
    $ 3266 "Home (Safe)"
    movej([-1.2302089344500047, -1.2969853503591224, -1.875639182904262, -1.539621866126728, 1.5731943360401213, -2.80099559440227], a=1.3962634015954636, v=1.0471975511965976)
  elif (45 == switch_1):
    $ 3267 "Case 45"
    $ 3268 "Place the decapped container- recipe"
    $ 3269 "tilt_to_home()"
    tilt_to_home()
    # begin: URCap Program Node
    #   Source: SensoPart VISOR Robotic, 2.0.6, SensoPart Industriesensorik GmbH
    #   Type: VISOR Robotic App
    $ 3271 "VISOR Easy Pick"
    def visorFuncEasyPick_fdc6d2():
      # begin: URCap Program Node
      #   Source: SensoPart VISOR Robotic, 2.0.6, SensoPart Industriesensorik GmbH
      #   Type: Easy Pick Setup
      $ 3272 "# 1 Setup" "noBreak"
      local easyPickVisorId = 1
      local easyPickArmMounted = True
      local easyPickSetJob = True
      local easyPickJobName = "PoTS"
      local easyPickAtImgAcq = False
      local easyPickImgAcqPose = Trigger
      # end: URCap Program Node
      # begin: URCap Program Node
      #   Source: SensoPart VISOR Robotic, 2.0.6, SensoPart Industriesensorik GmbH
      #   Type: Process
      $ 3273 "Process" "noBreak"
      local easyPickObjTaken = False
      local easyPickTrigger = False
      local easyPickPoseIdx = 0
      local easyPickPose = p[0,0,0,0,0,0]
      def easyPickFuncTrigger(visorId, setJob, jobName, arm):
      if (setJob):
        visor_changeJob(visorId, jobName, 6000)
      end
      if (arm):
        visor_trigger(visorId, 6000, "arm")
      else:
        visor_trigger(visorId, 6000)
      end
      global easyPickParts_7=visor_partsFound(visorId)
      visor_easyPickUpdate(visorId, "parts", visor_partsFound(visorId))
      return visor_getPose3d(visorId, 0)
    end
    while (not easyPickObjTaken):
      easyPickTrigger = (easyPickCount_7 >= visor_partsFound(easyPickVisorId)) or (easyPickCount_7 > 9) or (not visor_easyPickCheckIdent("d80e5c", easyPickVisorId))
      if (easyPickTrigger):
        easyPickCount_7 = 0
      end
      easyPickPoseIdx = easyPickCount_7
      easyPickPose = visor_getPose3d(easyPickVisorId, easyPickPoseIdx)
      visor_easyPickUpdate(easyPickVisorId, "counter", easyPickPoseIdx)
      # begin: URCap Program Node
      #   Source: SensoPart VISOR Robotic, 2.0.6, SensoPart Industriesensorik GmbH
      #   Type: Image Acquisition Pose
      $ 3274 "Image Acquisition Pose" "noBreak"
      if (easyPickTrigger):
        if (not easyPickAtImgAcq):
          movej(pose_trans(easyPickImgAcqPose,p[0.0000,0.0000,-0.0000,0.0000,0.0000,0.0000]),a=1.3963,v=1.0472,t=0.000000,r=0.000000)
          easyPickAtImgAcq = True
        end
        easyPickPose = easyPickFuncTrigger(easyPickVisorId, easyPickSetJob, easyPickJobName, easyPickArmMounted)
      end
      # end: URCap Program Node
      # begin: URCap Program Node
      #   Source: SensoPart VISOR Robotic, 2.0.6, SensoPart Industriesensorik GmbH
      #   Type: Object Detected
      $ 3275 "Object Detected" "noBreak"
      if (visor_partsFound(easyPickVisorId) > 0):
        $ 3276 "Open Gripper" "noBreak"
        # begin: URCap Program Node
        #   Source: Robotiq_Grippers, 3.17.0.105337, Robotiq Inc.
        #   Type: Gripper
        $ 3277 "Gripper Open (1)" "noBreak"
        if not(gripper_connected[0]):
          popup("Gripper 1 must be connected to run this program.", "No connection", False, True, True)
        end
        if not(rq_is_gripper_activated("1")):
          popup("Gripper 1 is not activated. Go to Installation tab > Gripper to activate it and run the program again.", "Not activated", False, True, True)
        end
        rq_set_pos_spd_for(0, 77, 77, "1")
        rq_wait_pos_spe_for_request(0, 77, 77, "1")
        rq_go_to("1")
        rq_wait("1")
        # end: URCap Program Node
        $ 3278 "Set" "noBreak"
        set_tcp(p[0.0,0.0,0.15052000000000001,3.1415,0.0,0.0])
        $ 3279 "Wait: 0.25" "noBreak"
        sleep(0.25)
        $ 3280 "MoveL" "noBreak"
        $ 3281 "OP_PowderA2" "noBreak"
        movel(OP_PowderA2_p, a=1.2, v=0.25)
        $ 3282 "Decap_up" "noBreak"
        movel(Decap_up_p, a=1.2, v=0.25)
        $ 3283 "Decap_pick" "noBreak"
        movel(Decap_pick_p, a=1.2, v=0.25)
        # begin: URCap Program Node
        #   Source: Robotiq_Grippers, 3.17.0.105337, Robotiq Inc.
        #   Type: Gripper
        $ 3284 "Gripper Close (1)" "noBreak"
        if not(gripper_connected[0]):
          popup("Gripper 1 must be connected to run this program.", "No connection", False, True, True)
        end
        if not(rq_is_gripper_activated("1")):
          popup("Gripper 1 is not activated. Go to Installation tab > Gripper to activate it and run the program again.", "Not activated", False, True, True)
        end
        rq_set_pos_spd_for(255, 77, 77, "1")
        rq_wait_pos_spe_for_request(255, 77, 77, "1")
        rq_go_to("1")
        rq_wait("1")
        # end: URCap Program Node
        $ 3285 "Wait: 0.5" "noBreak"
        sleep(0.5)
        $ 3286 "Set GRP_3F_Open=On" "noBreak"
        set_standard_digital_out(5, True)
        $ 3287 "Decap_up" "noBreak"
        movel(Decap_up_p, a=0.5, v=0.1)
        $ 3289 "Op_PowA_wP" "noBreak"
        movel(Op_PowA_wP_p, a=1.2, v=0.25)
        # begin: URCap Program Node
        #   Source: SensoPart VISOR Robotic, 2.0.6, SensoPart Industriesensorik GmbH
        #   Type: Approach Pose
        $ 3290 "Approach Pose" "noBreak"
        movej(pose_trans(easyPickPose,p[0.0000,0.0000,-0.0000,0.0000,0.0000,0.0000]),a=0.5236,v=0.4363,t=0.000000,r=0.000000)
        # end: URCap Program Node
        # begin: URCap Program Node
        #   Source: SensoPart VISOR Robotic, 2.0.6, SensoPart Industriesensorik GmbH
        #   Type: Target Pose
        $ 3291 "Target Pose" "noBreak"
        movel(pose_trans(easyPickPose,p[0.0000,0.0000,-0.0000,0.0000,0.0000,0.0000]),a=0.1000,v=0.0500,t=0.000000,r=0.000000)
        # end: URCap Program Node
        $ 3292 "Close Gripper" "noBreak"
        $ 3293 "container_place≔get_actual_tcp_pose()" "noBreak"
        global container_place= get_actual_tcp_pose ()
        $ 3294 "target_pose≔pose_add(container_place, p[0,0,-0.12,0,0,0])" "noBreak"
        global target_pose=pose_add(container_place, p[0,0,-0.12,0,0,0])
        $ 3295 "MoveL" "noBreak"
        $ 3296 "target_pose" "noBreak"
        movel(target_pose, a=0.3, v=0.05)
        # begin: URCap Program Node
        #   Source: Robotiq_Grippers, 3.17.0.105337, Robotiq Inc.
        #   Type: Gripper
        $ 3297 "Gripper Open (1)" "noBreak"
        if not(gripper_connected[0]):
          popup("Gripper 1 must be connected to run this program.", "No connection", False, True, True)
        end
        if not(rq_is_gripper_activated("1")):
          popup("Gripper 1 is not activated. Go to Installation tab > Gripper to activate it and run the program again.", "Not activated", False, True, True)
        end
        rq_set_pos_spd_for(0, 77, 77, "1")
        rq_wait_pos_spe_for_request(0, 77, 77, "1")
        rq_go_to("1")
        rq_wait("1")
        # end: URCap Program Node
        # begin: URCap Program Node
        #   Source: SensoPart VISOR Robotic, 2.0.6, SensoPart Industriesensorik GmbH
        #   Type: Exit Pose
        $ 3298 "Exit Pose" "noBreak"
        movel(pose_trans(easyPickPose,p[0.0000,0.0000,-0.0000,0.0000,0.0000,0.0000]),a=0.5000,v=0.2500,t=0.000000,r=0.000000)
        # end: URCap Program Node
        easyPickObjTaken = True
      end
      # end: URCap Program Node
      # begin: URCap Program Node
      #   Source: SensoPart VISOR Robotic, 2.0.6, SensoPart Industriesensorik GmbH
      #   Type: No Object Detected
      $ 3299 "No Object Detected" "noBreak"
      if (visor_partsFound(easyPickVisorId) < 1):
        $ 3300 "Popup: No weigh scale detected" "noBreak"
        popup("No weigh scale detected", "Message", False, False, blocking=True)
        else:
      end
      # end: URCap Program Node
    end
    easyPickCount_7 = easyPickCount_7 + 1
    visor_easyPickUpdate(easyPickVisorId, "counter", easyPickCount_7)
    visor_easyPickSetIdent("d80e5c", easyPickVisorId)
    # end: URCap Program Node
  end
  visorFuncEasyPick_fdc6d2()
  # end: URCap Program Node
  $ 3301 "place_pose≔get_actual_tcp_pose()"
  global place_pose= get_actual_tcp_pose ()
  $ 3302 "center_pose()"
  center_pose()
  $ 3304 "MoveJ"
  $ 3305 "Waypoint_1" "breakAfter"
  movej(get_inverse_kin(Waypoint_1_p, qnear=Waypoint_1_q), a=1.3962634015954636, v=1.0471975511965976)
  elif (46 == switch_1):
    $ 3306 "Case 46"
    $ 3307 "Powder dosing for recipe"
    $ 3309 "send_target_info()"
    send_target_info()
    $ 3310 "Wait: 0.5"
    sleep(0.5)
    $ 3311 "send_powder_info()"
    send_powder_info()
    $ 3312 "Wait: 0.5"
    sleep(0.5)
    # begin: URCap Program Node
    #   Source: SensoPart VISOR Robotic, 2.0.6, SensoPart Industriesensorik GmbH
    #   Type: VISOR Robotic App
    $ 3319 "VISOR Easy Pick"
    def visorFuncEasyPick_6dee13():
      # begin: URCap Program Node
      #   Source: SensoPart VISOR Robotic, 2.0.6, SensoPart Industriesensorik GmbH
      #   Type: Easy Pick Setup
      $ 3320 "# 1 Setup" "noBreak"
      local easyPickVisorId = 1
      local easyPickArmMounted = True
      local easyPickSetJob = True
      local easyPickJobName = "Weight_scale"
      local easyPickAtImgAcq = False
      local easyPickImgAcqPose = Trigger
      # end: URCap Program Node
      # begin: URCap Program Node
      #   Source: SensoPart VISOR Robotic, 2.0.6, SensoPart Industriesensorik GmbH
      #   Type: Process
      $ 3321 "Process" "noBreak"
      local easyPickObjTaken = False
      local easyPickTrigger = False
      local easyPickPoseIdx = 0
      local easyPickPose = p[0,0,0,0,0,0]
      def easyPickFuncTrigger(visorId, setJob, jobName, arm):
      if (setJob):
        visor_changeJob(visorId, jobName, 6000)
      end
      if (arm):
        visor_trigger(visorId, 6000, "arm")
      else:
        visor_trigger(visorId, 6000)
      end
      global easyPickParts_4=visor_partsFound(visorId)
      visor_easyPickUpdate(visorId, "parts", visor_partsFound(visorId))
      return visor_getPose3d(visorId, 0)
    end
    while (not easyPickObjTaken):
      easyPickTrigger = (easyPickCount_4 >= visor_partsFound(easyPickVisorId)) or (easyPickCount_4 > 9) or (not visor_easyPickCheckIdent("70b625", easyPickVisorId))
      if (easyPickTrigger):
        easyPickCount_4 = 0
      end
      easyPickPoseIdx = easyPickCount_4
      easyPickPose = visor_getPose3d(easyPickVisorId, easyPickPoseIdx)
      visor_easyPickUpdate(easyPickVisorId, "counter", easyPickPoseIdx)
      # begin: URCap Program Node
      #   Source: SensoPart VISOR Robotic, 2.0.6, SensoPart Industriesensorik GmbH
      #   Type: Image Acquisition Pose
      $ 3322 "Image Acquisition Pose" "noBreak"
      if (easyPickTrigger):
        if (not easyPickAtImgAcq):
          movej(pose_trans(easyPickImgAcqPose,p[0.0000,0.0000,-0.0000,0.0000,0.0000,0.0000]),a=1.3963,v=1.0472,t=0.000000,r=0.000000)
          easyPickAtImgAcq = True
        end
        easyPickPose = easyPickFuncTrigger(easyPickVisorId, easyPickSetJob, easyPickJobName, easyPickArmMounted)
      end
      # end: URCap Program Node
      # begin: URCap Program Node
      #   Source: SensoPart VISOR Robotic, 2.0.6, SensoPart Industriesensorik GmbH
      #   Type: Object Detected
      $ 3323 "Object Detected" "noBreak"
      if (visor_partsFound(easyPickVisorId) > 0):
        $ 3324 "Open Gripper" "noBreak"
        $ 3325 "tare_scale()" "noBreak"
        tare_scale()
        $ 3326 "Wait: 0.2" "noBreak"
        sleep(0.2)
        $ 3327 "weight_value≔get_weight()" "noBreak"
        global weight_value=get_weight()
        $ 3328 "Wait: 0.2" "noBreak"
        sleep(0.2)
        $ 3329 "diff≔target_weight-weight_value" "noBreak"
        global diff=target_weight-weight_value
        $ 3330 "scooping_init()" "noBreak"
        scooping_init()
        $ 3331 "compute_level_percent(W_now, weight_value)" "noBreak"
        compute_level_percent(W_now, weight_value)
        $ 3332 "send_level_info()" "noBreak"
        send_level_info()
        $ 3334 "spatula≔select_spatula(Flowability,level,diff,density)" "noBreak"
        global spatula=select_spatula(Flowability,level,diff,density)
        $ 3335 "Wait: 0.2" "noBreak"
        sleep(0.2)
        $ 3336 "send_spatula_info()" "noBreak"
        send_spatula_info()
        $ 3337 "If spatula ≟ 'spatula_L'" "noBreak"
        if (spatula  ==  "spatula_L"):
          $ 3338 "MoveJ" "noBreak"
          $ 3339 "Spatula_otw" "noBreak"
          movej(get_inverse_kin(Spatula_otw_p, qnear=Spatula_otw_q), a=1.3962634015954636, v=1.0471975511965976)
          $ 3340 "pick_spat_L_abv" "noBreak"
          movej(get_inverse_kin(pick_spat_L_abv_p, qnear=pick_spat_L_abv_q), a=1.3962634015954636, v=1.0471975511965976)
          $ 3341 "MoveL" "noBreak"
          $ 3342 "spat_L_pick" "noBreak"
          movel(spat_L_pick_p, a=1.2, v=0.25)
          # begin: URCap Program Node
          #   Source: Robotiq_Grippers, 3.17.0.105337, Robotiq Inc.
          #   Type: Gripper
          $ 3343 "Gripper Close (1)" "noBreak"
          if not(gripper_connected[0]):
            popup("Gripper 1 must be connected to run this program.", "No connection", False, True, True)
          end
          if not(rq_is_gripper_activated("1")):
            popup("Gripper 1 is not activated. Go to Installation tab > Gripper to activate it and run the program again.", "Not activated", False, True, True)
          end
          rq_set_pos_spd_for(255, 0, 77, "1")
          rq_wait_pos_spe_for_request(255, 0, 77, "1")
          rq_go_to("1")
          rq_wait("1")
          # end: URCap Program Node
          $ 3344 "spat_L_lift" "noBreak"
          movel(spat_L_lift_p, a=1.2, v=0.25, r=0.01)
          $ 3345 "spat_L_side" "noBreak"
          movel(spat_L_side_p, a=1.2, v=0.25, r=0.01)
          $ 3346 "spat_L_up" "noBreak"
          movel(spat_L_up_p, a=1.2, v=0.25, r=0.05)
          $ 3347 "MoveJ" "noBreak"
          $ 3348 "Spatula_otw" "noBreak"
          movej(get_inverse_kin(Spatula_otw_p, qnear=Spatula_otw_q), a=1.3962634015954636, v=1.0471975511965976)
        else:
          $ 3349 "ElseIf spatula ≟'spatula_M'" "noBreak"
          if (spatula  == "spatula_M"):
            $ 3350 "MoveJ" "noBreak"
            $ 3351 "Spatula_otw" "noBreak"
            movej(get_inverse_kin(Spatula_otw_p, qnear=Spatula_otw_q), a=1.3962634015954636, v=1.0471975511965976)
            $ 3352 "spat_M_up" "noBreak"
            movej(get_inverse_kin(spat_M_up_p, qnear=spat_M_up_q), a=1.3962634015954636, v=1.0471975511965976, r=0.05)
            $ 3353 "MoveL" "noBreak"
            $ 3354 "spat_M_pick" "noBreak"
            movel(spat_M_pick_p, a=1.2, v=0.25)
            # begin: URCap Program Node
            #   Source: Robotiq_Grippers, 3.17.0.105337, Robotiq Inc.
            #   Type: Gripper
            $ 3355 "Gripper Close (1)" "noBreak"
            if not(gripper_connected[0]):
              popup("Gripper 1 must be connected to run this program.", "No connection", False, True, True)
            end
            if not(rq_is_gripper_activated("1")):
              popup("Gripper 1 is not activated. Go to Installation tab > Gripper to activate it and run the program again.", "Not activated", False, True, True)
            end
            rq_set_pos_spd_for(255, 0, 77, "1")
            rq_wait_pos_spe_for_request(255, 0, 77, "1")
            rq_go_to("1")
            rq_wait("1")
            # end: URCap Program Node
            $ 3356 "spat_M_up" "noBreak"
            movel(spat_M_up_p, a=1.2, v=0.25, r=0.05)
            $ 3357 "Spatula_otw" "noBreak"
            movel(Spatula_otw_p, a=1.2, v=0.25)
            $ 3358 "switch_spat_M≔ False " "noBreak"
            global switch_spat_M=  False
          else:
            $ 3359 "ElseIf spatula≟'spatula_S'" "noBreak"
            if (spatula == "spatula_S"):
              $ 3360 "MoveJ" "noBreak"
              $ 3361 "Spatula_otw" "noBreak"
              movej(get_inverse_kin(Spatula_otw_p, qnear=Spatula_otw_q), a=1.3962634015954636, v=1.0471975511965976)
              $ 3362 "spat_S_Up_9" "noBreak"
              movej(get_inverse_kin(spat_S_Up_9_p, qnear=spat_S_Up_9_q), a=1.3962634015954636, v=1.0471975511965976, r=0.05)
              $ 3363 "MoveL" "noBreak"
              $ 3364 "spat_S_Pick_5" "noBreak"
              movel(spat_S_Pick_5_p, a=1.2, v=0.25)
              # begin: URCap Program Node
              #   Source: Robotiq_Grippers, 3.17.0.105337, Robotiq Inc.
              #   Type: Gripper
              $ 3365 "Gripper Close (1)" "noBreak"
              if not(gripper_connected[0]):
                popup("Gripper 1 must be connected to run this program.", "No connection", False, True, True)
              end
              if not(rq_is_gripper_activated("1")):
                popup("Gripper 1 is not activated. Go to Installation tab > Gripper to activate it and run the program again.", "Not activated", False, True, True)
              end
              rq_set_pos_spd_for(255, 0, 77, "1")
              rq_wait_pos_spe_for_request(255, 0, 77, "1")
              rq_go_to("1")
              rq_wait("1")
              # end: URCap Program Node
              $ 3366 "spat_S_Up_10" "noBreak"
              movel(spat_S_Up_10_p, a=1.2, v=0.25, r=0.05)
              $ 3367 "Spatula_otw" "noBreak"
              movel(Spatula_otw_p, a=1.2, v=0.25)
              $ 3368 "switch_spat_S≔ False " "noBreak"
              global switch_spat_S=  False
            else:
              $ 3369 "ElseIf spatula≟'spatula_flat_M'" "noBreak"
              if (spatula == "spatula_flat_M"):
                $ 3370 "MoveJ" "noBreak"
                $ 3371 "Spatula_otw" "noBreak"
                movej(get_inverse_kin(Spatula_otw_p, qnear=Spatula_otw_q), a=1.3962634015954636, v=1.0471975511965976)
                $ 3372 "spat_flatM_up" "noBreak"
                movej(get_inverse_kin(spat_flatM_up_p, qnear=spat_flatM_up_q), a=1.3962634015954636, v=1.0471975511965976, r=0.05)
                $ 3373 "MoveL" "noBreak"
                $ 3374 "spat_flatM_pick" "noBreak"
                movel(spat_flatM_pick_p, a=1.2, v=0.25)
                # begin: URCap Program Node
                #   Source: Robotiq_Grippers, 3.17.0.105337, Robotiq Inc.
                #   Type: Gripper
                $ 3375 "Gripper Close (1)" "noBreak"
                if not(gripper_connected[0]):
                  popup("Gripper 1 must be connected to run this program.", "No connection", False, True, True)
                end
                if not(rq_is_gripper_activated("1")):
                  popup("Gripper 1 is not activated. Go to Installation tab > Gripper to activate it and run the program again.", "Not activated", False, True, True)
                end
                rq_set_pos_spd_for(255, 0, 77, "1")
                rq_wait_pos_spe_for_request(255, 0, 77, "1")
                rq_go_to("1")
                rq_wait("1")
                # end: URCap Program Node
                $ 3376 "spat_flatM_up" "noBreak"
                movel(spat_flatM_up_p, a=1.2, v=0.25, r=0.05)
                $ 3377 "Spatula_otw" "noBreak"
                movel(Spatula_otw_p, a=1.2, v=0.25)
                $ 3378 "switch_spat_F_M≔ False " "noBreak"
                global switch_spat_F_M=  False
              else:
                $ 3379 "ElseIf spatula≟'spatula_flat_S'" "noBreak"
                if (spatula == "spatula_flat_S"):
                  $ 3380 "MoveJ" "noBreak"
                  $ 3381 "Spatula_otw" "noBreak"
                  movej(get_inverse_kin(Spatula_otw_p, qnear=Spatula_otw_q), a=1.3962634015954636, v=1.0471975511965976)
                  $ 3382 "spat_flatS_up" "noBreak"
                  movej(get_inverse_kin(spat_flatS_up_p, qnear=spat_flatS_up_q), a=1.3962634015954636, v=1.0471975511965976, r=0.05)
                  $ 3383 "MoveL" "noBreak"
                  $ 3384 "spat_flatS_pick" "noBreak"
                  movel(spat_flatS_pick_p, a=1.2, v=0.25)
                  # begin: URCap Program Node
                  #   Source: Robotiq_Grippers, 3.17.0.105337, Robotiq Inc.
                  #   Type: Gripper
                  $ 3385 "Gripper Close (1)" "noBreak"
                  if not(gripper_connected[0]):
                    popup("Gripper 1 must be connected to run this program.", "No connection", False, True, True)
                  end
                  if not(rq_is_gripper_activated("1")):
                    popup("Gripper 1 is not activated. Go to Installation tab > Gripper to activate it and run the program again.", "Not activated", False, True, True)
                  end
                  rq_set_pos_spd_for(255, 0, 77, "1")
                  rq_wait_pos_spe_for_request(255, 0, 77, "1")
                  rq_go_to("1")
                  rq_wait("1")
                  # end: URCap Program Node
                  $ 3386 "spat_flatS_up" "noBreak"
                  movel(spat_flatS_up_p, a=1.2, v=0.25, r=0.05)
                  $ 3387 "Spatula_otw" "noBreak"
                  movel(Spatula_otw_p, a=1.2, v=0.25)
                  $ 3388 "switch_spat_F_S≔ False " "noBreak"
                  global switch_spat_F_S=  False
                end
              end
            end
          end
        end
        $ 3389 "weight_value≔get_weight()" "noBreak"
        global weight_value=get_weight()
        $ 3390 "auto_tilt_and_scoop(W_now, target_weight, weight_value)" "noBreak"
        auto_tilt_and_scoop(W_now, target_weight, weight_value)
        # begin: URCap Program Node
        #   Source: SensoPart VISOR Robotic, 2.0.6, SensoPart Industriesensorik GmbH
        #   Type: Approach Pose
        $ 3391 "Approach Pose" "noBreak"
        movej(pose_trans(easyPickPose,p[0.0000,0.0000,0.0300,0.0000,0.0000,0.0000]),a=0.2618,v=0.1745,t=0.000000,r=0.000000)
        # end: URCap Program Node
        # begin: URCap Program Node
        #   Source: SensoPart VISOR Robotic, 2.0.6, SensoPart Industriesensorik GmbH
        #   Type: Target Pose
        $ 3392 "Target Pose" "noBreak"
        movel(pose_trans(easyPickPose,p[0.0000,0.0000,-0.0000,0.0000,0.0000,0.0000]),a=0.0500,v=0.0200,t=0.000000,r=0.000000)
        # end: URCap Program Node
        $ 3393 "Close Gripper" "noBreak"
        $ 3394 "dispense_pos≔get_actual_tcp_pose()" "noBreak"
        global dispense_pos= get_actual_tcp_pose ()
        $ 3395 "Loop weight_value≤target_weight" "noBreak"
        thread Thread_while_3395():
          while (True):
            $ 3396 "MoveL" "noBreak"
            $ 3397 "dispense_pos" "noBreak"
            movel(dispense_pos, a=0.2, v=0.1)
            $ 3398 "log_weight()" "noBreak"
            log_weight()
            $ 3399 "Wait: 0.5" "noBreak"
            sleep(0.5)
            $ 3400 "If level≥90.0" "noBreak"
            if (level >= 90.0):
              $ 3401 "Rotate()" "noBreak"
              Rotate()
            end
            $ 3402 "If level≤85" "noBreak"
            if (level <= 85):
              $ 3403 "tilt_to_home()" "noBreak"
              tilt_to_home()
            end
            $ 3404 "Wait: 0.5" "noBreak"
            sleep(0.5)
            $ 3405 "Start_thread≔ True " "noBreak"
            global Start_thread=  True
            $ 3406 "vib_thread≔ True " "noBreak"
            global vib_thread=  True
            $ 3408 "Wait: 0.5" "noBreak"
            sleep(0.5)
            $ 3414 "If diff ≥(target_g +(0.1*target_g))" "noBreak"
            if (diff  >= (target_g +(0.1*target_g))):
              $ 3415 "tilt_pose≔pose_trans(get_actual_tcp_pose(), p[0, 0, 0, 0, 0, 2.0])" "noBreak"
              global tilt_pose=pose_trans(get_actual_tcp_pose(), p[0, 0, 0, 0, 0, 2.0])
              $ 3416 "movel(tilt_pose, a=0.1, v=0.1, r=0.00001)" "noBreak"
              movel(tilt_pose, a=0.1, v=0.1, r=0.00001)
            else:
              $ 3417 "Else" "noBreak"
              $ 3418 "Loop weight_value≤target_weight and tilt_angle≥(-1.999) and tilt_angle≤0.5" "noBreak"
              thread Thread_while_3418():
                while (True):
                  $ 3419 "current_error≔target_weight-weight_value" "noBreak"
                  global current_error=target_weight-weight_value
                  $ 3420 "Integral_error≔Integral_error+current_error*dt" "noBreak"
                  global Integral_error=Integral_error+current_error*dt
                  $ 3421 "derivative≔(current_error-previous_error)/dt" "noBreak"
                  global derivative=(current_error-previous_error)/dt
                  $ 3422 "tilt_increment≔(kp*current_error)+(ki*Integral_error)+(kd*derivative)" "noBreak"
                  global tilt_increment=(kp*current_error)+(ki*Integral_error)+(kd*derivative)
                  $ 3423 "current_pose≔get_actual_tcp_pose()" "noBreak"
                  global current_pose= get_actual_tcp_pose ()
                  $ 3424 "tilt_angle≔current_pose[5]" "noBreak"
                  global tilt_angle=current_pose[5]
                  $ 3425 "tilt_pose≔pose_trans(current_pose, p[0, 0, 0, 0, 0, tilt_increment])" "noBreak"
                  global tilt_pose=pose_trans(current_pose, p[0, 0, 0, 0, 0, tilt_increment])
                  $ 3426 "movel(tilt_pose, a=0.1, v=0.1, r=0.00001)" "noBreak"
                  movel(tilt_pose, a=0.1, v=0.1, r=0.00001)
                  $ 3427 "previous_error≔current_error" "noBreak"
                  global previous_error=current_error
                end
              end
              if (weight_value <= target_weight  and  tilt_angle >= (-1.999)  and  tilt_angle <= 0.5):
                global thread_handler_3418=run Thread_while_3418()
                while (weight_value <= target_weight  and  tilt_angle >= (-1.999)  and  tilt_angle <= 0.5):
                  sync()
                end
                kill thread_handler_3418
              end
            end
            $ 3428 "Start_thread≔ False " "noBreak"
            global Start_thread=  False
            $ 3430 "weight_value≔get_weight()" "noBreak"
            global weight_value=get_weight()
            $ 3431 "tilt_angle≔-1" "noBreak"
            global tilt_angle=-1
            $ 3432 "Wait: 0.5" "noBreak"
            sleep(0.5)
            $ 3433 "vib_thread≔ False " "noBreak"
            global vib_thread=  False
            $ 3434 "MoveL" "noBreak"
            $ 3435 "dispense_pos" "noBreak"
            movel(dispense_pos, a=0.5, v=0.25)
            $ 3436 "compute_level_percent(W_now, weight_value)" "noBreak"
            compute_level_percent(W_now, weight_value)
            $ 3437 "send_level_info()" "noBreak"
            send_level_info()
            $ 3439 "spatula≔select_spatula(Flowability,level,diff,density)" "noBreak"
            global spatula=select_spatula(Flowability,level,diff,density)
            $ 3440 "Wait: 0.2" "noBreak"
            sleep(0.2)
            $ 3442 "Integral_error≔0" "noBreak"
            global Integral_error=0
            $ 3443 "current_error≔0" "noBreak"
            global current_error=0
            $ 3444 "previous_error≔0" "noBreak"
            global previous_error=0
            $ 3445 "Set AO[0]=0.0" "noBreak"
            set_standard_analog_out(0, 0.0)
            $ 3446 "Wait: 0.2" "noBreak"
            sleep(0.2)
            $ 3447 "send_spatula_info()" "noBreak"
            send_spatula_info()
            $ 3448 "If spatula ≟ 'spatula_M' and switch_spat_M≟ True " "noBreak"
            if (spatula  ==  "spatula_M"  and  switch_spat_M ==   True  ):
              $ 3449 "MoveJ" "noBreak"
              $ 3450 "Spatula_otw" "noBreak"
              movej(get_inverse_kin(Spatula_otw_p, qnear=Spatula_otw_q), a=1.3962634015954636, v=1.0471975511965976)
              $ 3451 "spat_L_up" "noBreak"
              movej(get_inverse_kin(spat_L_up_p, qnear=spat_L_up_q), a=1.3962634015954636, v=1.0471975511965976)
              $ 3452 "MoveL" "noBreak"
              $ 3453 "spat_L_side" "noBreak"
              movel(spat_L_side_p, a=1.2, v=0.25)
              $ 3454 "spat_L_lift" "noBreak"
              movel(spat_L_lift_p, a=1.2, v=0.25)
              $ 3455 "spat_L_pick" "noBreak"
              movel(spat_L_pick_p, a=1.2, v=0.25)
              # begin: URCap Program Node
              #   Source: Robotiq_Grippers, 3.17.0.105337, Robotiq Inc.
              #   Type: Gripper
              $ 3456 "Gripper Open (1)" "noBreak"
              if not(gripper_connected[0]):
                popup("Gripper 1 must be connected to run this program.", "No connection", False, True, True)
              end
              if not(rq_is_gripper_activated("1")):
                popup("Gripper 1 is not activated. Go to Installation tab > Gripper to activate it and run the program again.", "Not activated", False, True, True)
              end
              rq_set_pos_spd_for(0, 255, 77, "1")
              rq_wait_pos_spe_for_request(0, 255, 77, "1")
              rq_go_to("1")
              rq_wait("1")
              # end: URCap Program Node
              $ 3457 "spat_M_pick" "noBreak"
              movel(spat_M_pick_p, a=1.2, v=0.25)
              # begin: URCap Program Node
              #   Source: Robotiq_Grippers, 3.17.0.105337, Robotiq Inc.
              #   Type: Gripper
              $ 3458 "Gripper Close (1)" "noBreak"
              if not(gripper_connected[0]):
                popup("Gripper 1 must be connected to run this program.", "No connection", False, True, True)
              end
              if not(rq_is_gripper_activated("1")):
                popup("Gripper 1 is not activated. Go to Installation tab > Gripper to activate it and run the program again.", "Not activated", False, True, True)
              end
              rq_set_pos_spd_for(255, 0, 77, "1")
              rq_wait_pos_spe_for_request(255, 0, 77, "1")
              rq_go_to("1")
              rq_wait("1")
              # end: URCap Program Node
              $ 3459 "spat_M_up" "noBreak"
              movel(spat_M_up_p, a=1.2, v=0.25)
              $ 3460 "Spatula_otw" "noBreak"
              movel(Spatula_otw_p, a=1.2, v=0.25)
              $ 3461 "switch_spat_M≔ False " "noBreak"
              global switch_spat_M=  False
            else:
              $ 3462 "ElseIf spatula ≟ 'spatula_S' and switch_spat_S ≟ True " "noBreak"
              if (spatula  ==  "spatula_S" and switch_spat_S  ==   True  ):
                $ 3463 "MoveL" "noBreak"
                $ 3464 "Spatula_otw" "noBreak"
                movel(Spatula_otw_p, a=1.2, v=0.25)
                $ 3465 "spat_M_up" "noBreak"
                movel(spat_M_up_p, a=1.2, v=0.25)
                $ 3466 "spat_M_pick" "noBreak"
                movel(spat_M_pick_p, a=1.2, v=0.25)
                # begin: URCap Program Node
                #   Source: Robotiq_Grippers, 3.17.0.105337, Robotiq Inc.
                #   Type: Gripper
                $ 3467 "Gripper Open (1)" "noBreak"
                if not(gripper_connected[0]):
                  popup("Gripper 1 must be connected to run this program.", "No connection", False, True, True)
                end
                if not(rq_is_gripper_activated("1")):
                  popup("Gripper 1 is not activated. Go to Installation tab > Gripper to activate it and run the program again.", "Not activated", False, True, True)
                end
                rq_set_pos_spd_for(0, 255, 77, "1")
                rq_wait_pos_spe_for_request(0, 255, 77, "1")
                rq_go_to("1")
                rq_wait("1")
                # end: URCap Program Node
                $ 3468 "spat_S_pick" "noBreak"
                movel(spat_S_pick_p, a=1.2, v=0.25)
                # begin: URCap Program Node
                #   Source: Robotiq_Grippers, 3.17.0.105337, Robotiq Inc.
                #   Type: Gripper
                $ 3469 "Gripper Close (1)" "noBreak"
                if not(gripper_connected[0]):
                  popup("Gripper 1 must be connected to run this program.", "No connection", False, True, True)
                end
                if not(rq_is_gripper_activated("1")):
                  popup("Gripper 1 is not activated. Go to Installation tab > Gripper to activate it and run the program again.", "Not activated", False, True, True)
                end
                rq_set_pos_spd_for(255, 0, 77, "1")
                rq_wait_pos_spe_for_request(255, 0, 77, "1")
                rq_go_to("1")
                rq_wait("1")
                # end: URCap Program Node
                $ 3470 "spat_S_up" "noBreak"
                movel(spat_S_up_p, a=1.2, v=0.25)
                $ 3471 "Spatula_otw" "noBreak"
                movel(Spatula_otw_p, a=1.2, v=0.25)
                $ 3472 "switch_spat_S≔ False " "noBreak"
                global switch_spat_S=  False
              else:
                $ 3473 "ElseIf spatula≟'spatula_flat_S'  and switch_spat_F_S ≟ True " "noBreak"
                if (spatula == "spatula_flat_S"   and  switch_spat_F_S  ==   True  ):
                  $ 3474 "MoveL" "noBreak"
                  $ 3475 "Spatula_otw" "noBreak"
                  movel(Spatula_otw_p, a=1.2, v=0.25)
                  $ 3476 "spat_flatM_up" "noBreak"
                  movel(spat_flatM_up_p, a=1.2, v=0.25)
                  $ 3477 "spat_flatM_pick" "noBreak"
                  movel(spat_flatM_pick_p, a=1.2, v=0.25)
                  # begin: URCap Program Node
                  #   Source: Robotiq_Grippers, 3.17.0.105337, Robotiq Inc.
                  #   Type: Gripper
                  $ 3478 "Gripper Open (1)" "noBreak"
                  if not(gripper_connected[0]):
                    popup("Gripper 1 must be connected to run this program.", "No connection", False, True, True)
                  end
                  if not(rq_is_gripper_activated("1")):
                    popup("Gripper 1 is not activated. Go to Installation tab > Gripper to activate it and run the program again.", "Not activated", False, True, True)
                  end
                  rq_set_pos_spd_for(0, 0, 77, "1")
                  rq_wait_pos_spe_for_request(0, 0, 77, "1")
                  rq_go_to("1")
                  rq_wait("1")
                  # end: URCap Program Node
                  $ 3479 "spat_flatS_pick" "noBreak"
                  movel(spat_flatS_pick_p, a=1.2, v=0.25)
                  # begin: URCap Program Node
                  #   Source: Robotiq_Grippers, 3.17.0.105337, Robotiq Inc.
                  #   Type: Gripper
                  $ 3480 "Gripper Close (1)" "noBreak"
                  if not(gripper_connected[0]):
                    popup("Gripper 1 must be connected to run this program.", "No connection", False, True, True)
                  end
                  if not(rq_is_gripper_activated("1")):
                    popup("Gripper 1 is not activated. Go to Installation tab > Gripper to activate it and run the program again.", "Not activated", False, True, True)
                  end
                  rq_set_pos_spd_for(255, 0, 77, "1")
                  rq_wait_pos_spe_for_request(255, 0, 77, "1")
                  rq_go_to("1")
                  rq_wait("1")
                  # end: URCap Program Node
                  $ 3481 "spat_flatS_up" "noBreak"
                  movel(spat_flatS_up_p, a=1.2, v=0.25)
                  $ 3482 "Spatula_otw" "noBreak"
                  movel(Spatula_otw_p, a=1.2, v=0.25)
                  $ 3483 "switch_spat_F_S≔ False " "noBreak"
                  global switch_spat_F_S=  False
                end
              end
            end
            $ 3484 "auto_tilt_and_scoop(W_now, target_weight, weight_value)" "noBreak"
            auto_tilt_and_scoop(W_now, target_weight, weight_value)
            $ 3485 "Wait: 0.5" "noBreak"
            sleep(0.5)
          end
        end
        if (weight_value <= target_weight):
          global thread_handler_3395=run Thread_while_3395()
          while (weight_value <= target_weight):
            sync()
          end
          kill thread_handler_3395
        end
        $ 3486 "Start_thread≔ False " "noBreak"
        global Start_thread=  False
        $ 3487 "Wait: 0.5" "noBreak"
        sleep(0.5)
        $ 3488 "vib_thread≔ False " "noBreak"
        global vib_thread=  False
        # begin: URCap Program Node
        #   Source: SensoPart VISOR Robotic, 2.0.6, SensoPart Industriesensorik GmbH
        #   Type: Exit Pose
        $ 3490 "Exit Pose" "noBreak"
        movel(pose_trans(easyPickPose,p[0.0000,0.0000,-0.0000,0.0000,0.0000,0.0000]),a=0.5000,v=0.2500,t=0.000000,r=0.000000)
        # end: URCap Program Node
        easyPickObjTaken = True
      end
      # end: URCap Program Node
      # begin: URCap Program Node
      #   Source: SensoPart VISOR Robotic, 2.0.6, SensoPart Industriesensorik GmbH
      #   Type: No Object Detected
      $ 3491 "No Object Detected" "noBreak"
      if (visor_partsFound(easyPickVisorId) < 1):
        $ 3492 "Popup: No weigh scale detected" "noBreak"
        popup("No weigh scale detected", "Message", False, False, blocking=True)
        else:
      end
      # end: URCap Program Node
    end
    easyPickCount_4 = easyPickCount_4 + 1
    visor_easyPickUpdate(easyPickVisorId, "counter", easyPickCount_4)
    visor_easyPickSetIdent("70b625", easyPickVisorId)
    # end: URCap Program Node
  end
  visorFuncEasyPick_6dee13()
  # end: URCap Program Node
  $ 3495 "MoveJ"
  $ 3496 "dispense_pos" "breakAfter"
  movej(dispense_pos, a=0.5235987755982988, v=0.4363323129985824)
  $ 3497 "weight_value≔get_weight()"
  global weight_value=get_weight()
  $ 3498 "after_scoop()"
  after_scoop()
  $ 3499 "Place spatula back to the rack"
  $ 3500 "If spatula≟'spatula_M'"
  if (spatula == "spatula_M"):
    $ 3501 "MoveJ"
    $ 3502 "Spatula_otw" "breakAfter"
    movej(get_inverse_kin(Spatula_otw_p, qnear=Spatula_otw_q), a=1.3962634015954636, v=1.0471975511965976)
    $ 3503 "spat_M_up" "breakAfter"
    movej(get_inverse_kin(spat_M_up_p, qnear=spat_M_up_q), a=1.3962634015954636, v=1.0471975511965976)
    $ 3504 "MoveL"
    $ 3505 "spat_M_pick" "breakAfter"
    movel(spat_M_pick_p, a=1.2, v=0.25)
    # begin: URCap Program Node
    #   Source: Robotiq_Grippers, 3.17.0.105337, Robotiq Inc.
    #   Type: Gripper
    $ 3506 "Gripper Open (1)"
    if not(gripper_connected[0]):
      popup("Gripper 1 must be connected to run this program.", "No connection", False, True, True)
    end
    if not(rq_is_gripper_activated("1")):
      popup("Gripper 1 is not activated. Go to Installation tab > Gripper to activate it and run the program again.", "Not activated", False, True, True)
    end
    rq_set_pos_spd_for(0, 128, 77, "1")
    rq_wait_pos_spe_for_request(0, 128, 77, "1")
    rq_go_to("1")
    rq_wait("1")
    # end: URCap Program Node
    $ 3507 "spat_M_up" "breakAfter"
    movel(spat_M_up_p, a=1.2, v=0.25)
    $ 3508 "Home (Safe)"
    movej([-1.2302089344500047, -1.2969853503591224, -1.875639182904262, -1.539621866126728, 1.5731943360401213, -2.80099559440227], a=1.3962634015954636, v=1.0471975511965976)
  else:
    $ 3509 "ElseIf spatula≟'spatula_flat_S'"
    if (spatula == "spatula_flat_S"):
      $ 3510 "MoveJ"
      $ 3511 "Spatula_otw" "breakAfter"
      movej(get_inverse_kin(Spatula_otw_p, qnear=Spatula_otw_q), a=1.3962634015954636, v=1.0471975511965976)
      $ 3512 "spat_flatS_up" "breakAfter"
      movej(get_inverse_kin(spat_flatS_up_p, qnear=spat_flatS_up_q), a=1.3962634015954636, v=1.0471975511965976)
      $ 3513 "MoveL"
      $ 3514 "spat_flatS_pick" "breakAfter"
      movel(spat_flatS_pick_p, a=1.2, v=0.25)
      # begin: URCap Program Node
      #   Source: Robotiq_Grippers, 3.17.0.105337, Robotiq Inc.
      #   Type: Gripper
      $ 3515 "Gripper Open (1)"
      if not(gripper_connected[0]):
        popup("Gripper 1 must be connected to run this program.", "No connection", False, True, True)
      end
      if not(rq_is_gripper_activated("1")):
        popup("Gripper 1 is not activated. Go to Installation tab > Gripper to activate it and run the program again.", "Not activated", False, True, True)
      end
      rq_set_pos_spd_for(0, 128, 77, "1")
      rq_wait_pos_spe_for_request(0, 128, 77, "1")
      rq_go_to("1")
      rq_wait("1")
      # end: URCap Program Node
      $ 3516 "spat_flatS_up" "breakAfter"
      movel(spat_flatS_up_p, a=1.2, v=0.25)
      $ 3517 "Home (Safe)"
      movej([-1.2302089344500047, -1.2969853503591224, -1.875639182904262, -1.539621866126728, 1.5731943360401213, -2.80099559440227], a=1.3962634015954636, v=1.0471975511965976)
    end
  end
  $ 3518 "Pick container from PoTS"
  $ 3519 "cont_place_offs≔pose_add(container_place, p[0.05,0,0,0,0,0])"
  global cont_place_offs=pose_add(container_place, p[0.05,0,0,0,0,0])
  $ 3520 "MoveJ"
  $ 3521 "cont_place_offs" "breakAfter"
  movej(cont_place_offs, a=1.3962634015954636, v=1.0471975511965976)
  $ 3522 "container_place" "breakAfter"
  movej(container_place, a=1.3962634015954636, v=1.0471975511965976)
  $ 3523 "MoveL"
  $ 3524 "target_pose" "breakAfter"
  movel(target_pose, a=1.2, v=0.25)
  # begin: URCap Program Node
  #   Source: Robotiq_Grippers, 3.17.0.105337, Robotiq Inc.
  #   Type: Gripper
  $ 3525 "Gripper Close (1)"
  if not(gripper_connected[0]):
    popup("Gripper 1 must be connected to run this program.", "No connection", False, True, True)
  end
  if not(rq_is_gripper_activated("1")):
    popup("Gripper 1 is not activated. Go to Installation tab > Gripper to activate it and run the program again.", "Not activated", False, True, True)
  end
  rq_set_pos_spd_for(255, 77, 77, "1")
  rq_wait_pos_spe_for_request(255, 77, 77, "1")
  rq_go_to("1")
  rq_wait("1")
  # end: URCap Program Node
  $ 3526 "container_place" "breakAfter"
  movel(container_place, a=0.6, v=0.1)
  $ 3528 "Place Powder container back to holder"
  $ 3529 "If powder_position ≟ 'Position1'"
  if (powder_position  ==  "Position1"):
    $ 3530 "MoveL"
    $ 3531 "Postions_otw" "breakAfter"
    movel(Postions_otw_p, a=1.2, v=0.25, r=0.01)
    $ 3532 "MoveL"
    $ 3533 "PosA_up" "breakAfter"
    movel(PosA_up_p, a=1.2, v=0.25)
    $ 3534 "PosA_pick" "breakAfter"
    movel(PosA_pick_p, a=0.3, v=0.05)
    # begin: URCap Program Node
    #   Source: Robotiq_Grippers, 3.17.0.105337, Robotiq Inc.
    #   Type: Gripper
    $ 3535 "Gripper Open (1)"
    if not(gripper_connected[0]):
      popup("Gripper 1 must be connected to run this program.", "No connection", False, True, True)
    end
    if not(rq_is_gripper_activated("1")):
      popup("Gripper 1 is not activated. Go to Installation tab > Gripper to activate it and run the program again.", "Not activated", False, True, True)
    end
    rq_set_pos_spd_for(0, 128, 77, "1")
    rq_wait_pos_spe_for_request(0, 128, 77, "1")
    rq_go_to("1")
    rq_wait("1")
    # end: URCap Program Node
    $ 3536 "PosA_up" "breakAfter"
    movel(PosA_up_p, a=1.2, v=0.25)
    $ 3537 "Postions_otw" "breakAfter"
    movel(Postions_otw_p, a=1.2, v=0.25, r=0.05)
  else:
    $ 3538 "ElseIf powder_position≟'Position2'"
    if (powder_position == "Position2"):
      $ 3539 "MoveL"
      $ 3540 "Postions_otw" "breakAfter"
      movel(Postions_otw_p, a=1.2, v=0.25, r=0.01)
      $ 3541 "MoveL"
      $ 3542 "PosB_up" "breakAfter"
      movel(PosB_up_p, a=1.2, v=0.25, r=0.01)
      $ 3543 "PosB_pick" "breakAfter"
      movel(PosB_pick_p, a=0.3, v=0.05)
      # begin: URCap Program Node
      #   Source: Robotiq_Grippers, 3.17.0.105337, Robotiq Inc.
      #   Type: Gripper
      $ 3544 "Gripper Open (1)"
      if not(gripper_connected[0]):
        popup("Gripper 1 must be connected to run this program.", "No connection", False, True, True)
      end
      if not(rq_is_gripper_activated("1")):
        popup("Gripper 1 is not activated. Go to Installation tab > Gripper to activate it and run the program again.", "Not activated", False, True, True)
      end
      rq_set_pos_spd_for(0, 128, 77, "1")
      rq_wait_pos_spe_for_request(0, 128, 77, "1")
      rq_go_to("1")
      rq_wait("1")
      # end: URCap Program Node
      $ 3545 "PosB_up" "breakAfter"
      movel(PosB_up_p, a=1.2, v=0.25)
      $ 3546 "Postions_otw" "breakAfter"
      movel(Postions_otw_p, a=1.2, v=0.25, r=0.05)
    else:
      $ 3547 "ElseIf powder_position≟'Position3'"
      if (powder_position == "Position3"):
        $ 3548 "MoveL"
        $ 3549 "Postions_otw" "breakAfter"
        movel(Postions_otw_p, a=1.2, v=0.25, r=0.01)
        $ 3550 "MoveL"
        $ 3551 "PosC_up" "breakAfter"
        movel(PosC_up_p, a=1.2, v=0.25, r=0.01)
        $ 3552 "PosC_pick" "breakAfter"
        movel(PosC_pick_p, a=0.3, v=0.05)
        # begin: URCap Program Node
        #   Source: Robotiq_Grippers, 3.17.0.105337, Robotiq Inc.
        #   Type: Gripper
        $ 3553 "Gripper Open (1)"
        if not(gripper_connected[0]):
          popup("Gripper 1 must be connected to run this program.", "No connection", False, True, True)
        end
        if not(rq_is_gripper_activated("1")):
          popup("Gripper 1 is not activated. Go to Installation tab > Gripper to activate it and run the program again.", "Not activated", False, True, True)
        end
        rq_set_pos_spd_for(0, 128, 77, "1")
        rq_wait_pos_spe_for_request(0, 128, 77, "1")
        rq_go_to("1")
        rq_wait("1")
        # end: URCap Program Node
        $ 3554 "PosC_up" "breakAfter"
        movel(PosC_up_p, a=1.2, v=0.25)
        $ 3555 "Postions_otw" "breakAfter"
        movel(Postions_otw_p, a=1.2, v=0.25, r=0.05)
      end
    end
  end
  $ 3556 "MoveJ"
  $ 3557 "Cap_above" "breakAfter"
  movej(get_inverse_kin(Cap_above_p, qnear=Cap_above_q), a=1.3962634015954636, v=1.0471975511965976, r=0.05)
  $ 3558 "MoveL"
  $ 3559 "Cap_place" "breakAfter"
  movel(Cap_place_p, a=1.2, v=0.25)
  # begin: URCap Program Node
  #   Source: Robotiq_Grippers, 3.17.0.105337, Robotiq Inc.
  #   Type: Gripper
  $ 3560 "Gripper Close (1)"
  if not(gripper_connected[0]):
    popup("Gripper 1 must be connected to run this program.", "No connection", False, True, True)
  end
  if not(rq_is_gripper_activated("1")):
    popup("Gripper 1 is not activated. Go to Installation tab > Gripper to activate it and run the program again.", "Not activated", False, True, True)
  end
  rq_set_pos_spd_for(255, 77, 77, "1")
  rq_wait_pos_spe_for_request(255, 77, 77, "1")
  rq_go_to("1")
  rq_wait("1")
  # end: URCap Program Node
  $ 3561 "Cap_above" "breakAfter"
  movel(Cap_above_p, a=1.2, v=0.25, r=0.05)
  $ 3562 "Cap the container"
  $ 3563 "If powder_position ≟ 'Position1'"
  if (powder_position  ==  "Position1"):
    $ 3564 "MoveJ"
    $ 3565 "Cap_Pos1_up" "breakAfter"
    movej(get_inverse_kin(Cap_Pos1_up_p, qnear=Cap_Pos1_up_q), a=1.3962634015954636, v=1.0471975511965976)
    $ 3566 "MoveL"
    $ 3567 "Cap_pos1" "breakAfter"
    movel(Cap_pos1_p, a=0.3, v=0.05)
  else:
    $ 3568 "ElseIf powder_position≟'Position2'"
    if (powder_position == "Position2"):
      $ 3569 "MoveJ"
      $ 3570 "Cap_Pos2_up" "breakAfter"
      movej(get_inverse_kin(Cap_Pos2_up_p, qnear=Cap_Pos2_up_q), a=1.3962634015954636, v=1.0471975511965976)
      $ 3571 "MoveL"
      $ 3572 "Cap_Pos2" "breakAfter"
      movel(Cap_Pos2_p, a=0.3, v=0.05)
    else:
      $ 3573 "ElseIf powder_position≟'Position3'"
      if (powder_position == "Position3"):
        $ 3574 "MoveJ"
        $ 3575 "Cap_Pos3_up" "breakAfter"
        movej(get_inverse_kin(Cap_Pos3_up_p, qnear=Cap_Pos3_up_q), a=1.3962634015954636, v=1.0471975511965976)
        $ 3576 "MoveL"
        $ 3577 "Cap_pos3" "breakAfter"
        movel(Cap_pos3_p, a=0.3, v=0.05)
      end
    end
  end
  $ 3578 "Capping motion"
  # begin: URCap Program Node
  #   Source: Robotiq_Grippers, 3.17.0.105337, Robotiq Inc.
  #   Type: Gripper
  $ 3579 "Gripper Move30mm (1)"
  if not(gripper_connected[0]):
    popup("Gripper 1 must be connected to run this program.", "No connection", False, True, True)
  end
  if not(rq_is_gripper_activated("1")):
    popup("Gripper 1 is not activated. Go to Installation tab > Gripper to activate it and run the program again.", "Not activated", False, True, True)
  end
  rq_set_pos_spd_for(110, 77, 77, "1")
  rq_wait_pos_spe_for_request(110, 77, 77, "1")
  rq_go_to("1")
  rq_wait("1")
  # end: URCap Program Node
  $ 3580 "Loop 2 times"
  Loop_7 = 0
  while (Loop_7 < 2):
    $ 3586 "Cap_CW≔pose_add(get_actual_tcp_pose(), p[0,0,0,0,0,2.2])"
    global Cap_CW= pose_add ( get_actual_tcp_pose (), p[0,0,0,0,0,2.2])
    $ 3587 "MoveL"
    $ 3588 "Cap_CW" "breakAfter"
    movel(Cap_CW, a=1.2, v=0.25)
    # begin: URCap Program Node
    #   Source: Robotiq_Grippers, 3.17.0.105337, Robotiq Inc.
    #   Type: Gripper
    $ 3589 "Gripper Move25mm (1)"
    if not(gripper_connected[0]):
      popup("Gripper 1 must be connected to run this program.", "No connection", False, True, True)
    end
    if not(rq_is_gripper_activated("1")):
      popup("Gripper 1 is not activated. Go to Installation tab > Gripper to activate it and run the program again.", "Not activated", False, True, True)
    end
    rq_set_pos_spd_for(133, 77, 77, "1")
    rq_wait_pos_spe_for_request(133, 77, 77, "1")
    rq_go_to("1")
    rq_wait("1")
    # end: URCap Program Node
    $ 3590 "Cap_CCW≔pose_add(get_actual_tcp_pose(), p[0,0,0,0,0,-2.2])"
    global Cap_CCW= pose_add ( get_actual_tcp_pose (), p[0,0,0,0,0,-2.2])
    $ 3591 "MoveL"
    $ 3592 "Cap_CCW" "breakAfter"
    movel(Cap_CCW, a=1.2, v=0.25)
    # begin: URCap Program Node
    #   Source: Robotiq_Grippers, 3.17.0.105337, Robotiq Inc.
    #   Type: Gripper
    $ 3593 "Gripper Move30mm (1)"
    if not(gripper_connected[0]):
      popup("Gripper 1 must be connected to run this program.", "No connection", False, True, True)
    end
    if not(rq_is_gripper_activated("1")):
      popup("Gripper 1 is not activated. Go to Installation tab > Gripper to activate it and run the program again.", "Not activated", False, True, True)
    end
    rq_set_pos_spd_for(110, 77, 77, "1")
    rq_wait_pos_spe_for_request(110, 77, 77, "1")
    rq_go_to("1")
    rq_wait("1")
    # end: URCap Program Node
    Loop_7 = Loop_7 + 1
  end
  # begin: URCap Program Node
  #   Source: Robotiq_Grippers, 3.17.0.105337, Robotiq Inc.
  #   Type: Gripper
  $ 3594 "Gripper Open (1)"
  if not(gripper_connected[0]):
    popup("Gripper 1 must be connected to run this program.", "No connection", False, True, True)
  end
  if not(rq_is_gripper_activated("1")):
    popup("Gripper 1 is not activated. Go to Installation tab > Gripper to activate it and run the program again.", "Not activated", False, True, True)
  end
  rq_set_pos_spd_for(0, 77, 77, "1")
  rq_wait_pos_spe_for_request(0, 77, 77, "1")
  rq_go_to("1")
  rq_wait("1")
  # end: URCap Program Node
  $ 3595 "after_capping≔pose_add(get_actual_tcp_pose(), p[0,0,0.05,0,0,0])"
  global after_capping=pose_add(get_actual_tcp_pose(), p[0,0,0.05,0,0,0])
  $ 3596 "MoveL"
  $ 3597 "after_capping" "breakAfter"
  movel(after_capping, a=1.2, v=0.25)
  $ 3598 "Home (Safe)"
  movej([-1.2302089344500047, -1.2969853503591224, -1.875639182904262, -1.539621866126728, 1.5731943360401213, -2.80099559440227], a=1.3962634015954636, v=1.0471975511965976)
  elif (47 == switch_1):
    $ 3599 "Case 47"
    $ 3600 "Pick containers"
    # begin: URCap Program Node
    #   Source: SensoPart VISOR Robotic, 2.0.6, SensoPart Industriesensorik GmbH
    #   Type: VISOR Robotic App
    $ 3601 "VISOR Easy Pick"
    def visorFuncEasyPick_c5f2c2():
      # begin: URCap Program Node
      #   Source: SensoPart VISOR Robotic, 2.0.6, SensoPart Industriesensorik GmbH
      #   Type: Easy Pick Setup
      $ 3602 "# 1 Setup" "noBreak"
      local easyPickVisorId = 1
      local easyPickArmMounted = True
      local easyPickSetJob = True
      local easyPickJobName = "Containers_pick"
      local easyPickAtImgAcq = False
      local easyPickImgAcqPose = Trigger
      # end: URCap Program Node
      # begin: URCap Program Node
      #   Source: SensoPart VISOR Robotic, 2.0.6, SensoPart Industriesensorik GmbH
      #   Type: Process
      $ 3603 "Process" "noBreak"
      local easyPickObjTaken = False
      local easyPickTrigger = False
      local easyPickPoseIdx = 0
      local easyPickPose = p[0,0,0,0,0,0]
      def easyPickFuncTrigger(visorId, setJob, jobName, arm):
      if (setJob):
        visor_changeJob(visorId, jobName, 6000)
      end
      if (arm):
        visor_trigger(visorId, 6000, "arm")
      else:
        visor_trigger(visorId, 6000)
      end
      global easyPickParts_9=visor_partsFound(visorId)
      visor_easyPickUpdate(visorId, "parts", visor_partsFound(visorId))
      return visor_getPose3d(visorId, 0)
    end
    while (not easyPickObjTaken):
      easyPickTrigger = (easyPickCount_9 >= visor_partsFound(easyPickVisorId)) or (easyPickCount_9 > 9) or (not visor_easyPickCheckIdent("b42f27", easyPickVisorId))
      if (easyPickTrigger):
        easyPickCount_9 = 0
      end
      easyPickPoseIdx = easyPickCount_9
      easyPickPose = visor_getPose3d(easyPickVisorId, easyPickPoseIdx)
      visor_easyPickUpdate(easyPickVisorId, "counter", easyPickPoseIdx)
      # begin: URCap Program Node
      #   Source: SensoPart VISOR Robotic, 2.0.6, SensoPart Industriesensorik GmbH
      #   Type: Image Acquisition Pose
      $ 3604 "Image Acquisition Pose" "noBreak"
      if (easyPickTrigger):
        if (not easyPickAtImgAcq):
          movej(pose_trans(easyPickImgAcqPose,p[0.0000,0.0000,-0.0000,0.0000,0.0000,0.0000]),a=1.3963,v=1.0472,t=0.000000,r=0.000000)
          easyPickAtImgAcq = True
        end
        easyPickPose = easyPickFuncTrigger(easyPickVisorId, easyPickSetJob, easyPickJobName, easyPickArmMounted)
      end
      # end: URCap Program Node
      # begin: URCap Program Node
      #   Source: SensoPart VISOR Robotic, 2.0.6, SensoPart Industriesensorik GmbH
      #   Type: Object Detected
      $ 3605 "Object Detected" "noBreak"
      if (visor_partsFound(easyPickVisorId) > 0):
        $ 3606 "Open Gripper" "noBreak"
        # begin: URCap Program Node
        #   Source: Robotiq_Grippers, 3.17.0.105337, Robotiq Inc.
        #   Type: Gripper
        $ 3607 "Gripper Open (1)" "noBreak"
        if not(gripper_connected[0]):
          popup("Gripper 1 must be connected to run this program.", "No connection", False, True, True)
        end
        if not(rq_is_gripper_activated("1")):
          popup("Gripper 1 is not activated. Go to Installation tab > Gripper to activate it and run the program again.", "Not activated", False, True, True)
        end
        rq_set_pos_spd_for(0, 77, 77, "1")
        rq_wait_pos_spe_for_request(0, 77, 77, "1")
        rq_go_to("1")
        rq_wait("1")
        # end: URCap Program Node
        $ 3608 "MoveJ" "noBreak"
        $ 3609 "pick_cont_otw" "noBreak"
        movej(get_inverse_kin(pick_cont_otw_p, qnear=pick_cont_otw_q), a=1.3962634015954636, v=1.0471975511965976)
        # begin: URCap Program Node
        #   Source: SensoPart VISOR Robotic, 2.0.6, SensoPart Industriesensorik GmbH
        #   Type: Approach Pose
        $ 3610 "Approach Pose" "noBreak"
        movej(pose_trans(easyPickPose,p[0.0000,0.0000,0.0500,0.0000,0.0000,0.0000]),a=1.3963,v=1.0472,t=0.000000,r=0.000000)
        # end: URCap Program Node
        # begin: URCap Program Node
        #   Source: SensoPart VISOR Robotic, 2.0.6, SensoPart Industriesensorik GmbH
        #   Type: Target Pose
        $ 3611 "Target Pose" "noBreak"
        movej(pose_trans(easyPickPose,p[0.0000,0.0000,-0.0000,0.0000,0.0000,0.0000]),a=1.3963,v=1.0472,t=0.000000,r=0.000000)
        # end: URCap Program Node
        $ 3612 "Close Gripper" "noBreak"
        # begin: URCap Program Node
        #   Source: Robotiq_Grippers, 3.17.0.105337, Robotiq Inc.
        #   Type: Gripper
        $ 3613 "Gripper Close (1)" "noBreak"
        if not(gripper_connected[0]):
          popup("Gripper 1 must be connected to run this program.", "No connection", False, True, True)
        end
        if not(rq_is_gripper_activated("1")):
          popup("Gripper 1 is not activated. Go to Installation tab > Gripper to activate it and run the program again.", "Not activated", False, True, True)
        end
        rq_set_pos_spd_for(255, 77, 77, "1")
        rq_wait_pos_spe_for_request(255, 77, 77, "1")
        rq_go_to("1")
        rq_wait("1")
        # end: URCap Program Node
        # begin: URCap Program Node
        #   Source: SensoPart VISOR Robotic, 2.0.6, SensoPart Industriesensorik GmbH
        #   Type: Exit Pose
        $ 3614 "Exit Pose" "noBreak"
        movej(pose_trans(easyPickPose,p[0.0000,0.0000,-0.0000,0.0000,0.0000,0.0000]),a=1.3963,v=1.0472,t=0.000000,r=0.000000)
        # end: URCap Program Node
        easyPickObjTaken = True
      end
      # end: URCap Program Node
      # begin: URCap Program Node
      #   Source: SensoPart VISOR Robotic, 2.0.6, SensoPart Industriesensorik GmbH
      #   Type: No Object Detected
      $ 3615 "No Object Detected" "noBreak"
      if (visor_partsFound(easyPickVisorId) < 1):
        $ 3616 "Popup: No container detected" "noBreak"
        popup("No container detected", "Message", False, False, blocking=True)
        else:
      end
      # end: URCap Program Node
    end
    easyPickCount_9 = easyPickCount_9 + 1
    visor_easyPickUpdate(easyPickVisorId, "counter", easyPickCount_9)
    visor_easyPickSetIdent("b42f27", easyPickVisorId)
    # end: URCap Program Node
  end
  visorFuncEasyPick_c5f2c2()
  # end: URCap Program Node
  $ 3617 "MoveJ"
  $ 3618 "Powder_wayp1" "breakAfter"
  movej(get_inverse_kin(Powder_wayp1_p, qnear=Powder_wayp1_q), a=1.3962634015954636, v=1.0471975511965976)
  $ 3619 "If powder_position ≟ 'Position1'"
  if (powder_position  ==  "Position1"):
    $ 3620 "MoveJ"
    $ 3621 "Postions_otw" "breakAfter"
    movej(get_inverse_kin(Postions_otw_p, qnear=Postions_otw_q), a=1.3962634015954636, v=1.0471975511965976, r=0.01)
    $ 3622 "MoveL"
    $ 3623 "PosA_up" "breakAfter"
    movel(PosA_up_p, a=1.2, v=0.25)
    $ 3624 "PosA_pick" "breakAfter"
    movel(PosA_pick_p, a=0.3, v=0.05)
    # begin: URCap Program Node
    #   Source: Robotiq_Grippers, 3.17.0.105337, Robotiq Inc.
    #   Type: Gripper
    $ 3625 "Gripper Open (1)"
    if not(gripper_connected[0]):
      popup("Gripper 1 must be connected to run this program.", "No connection", False, True, True)
    end
    if not(rq_is_gripper_activated("1")):
